REGION Network 36: STATE Num:120 StNextRdyInTransit
   RUNG wire#powerrail
      Contact( #sStNextRdyInTransit )
      wire#w1
      I_Contact( #sStWtResetRel )
      I_Contact( #sStNextRdyInTransit_T1 )
      I_Contact( #sStNextRdyInTransit_T2 )
      wire#w2
      Coil( #sStNextRdyInTransit )
   END_RUNG
   RUNG wire#powerrail
      Contact( #sStRecovery_T4 )
   END_RUNG wire#w1
   RUNG wire#powerrail
      Contact( #sStWtLifterAtPosn1_T1 )
   END_RUNG wire#w1
   RUNG wire#w2
      { S7_GenerateENO := "TRUE" } Move(in := 120, out1 => #StateNo)
   END_RUNG
   // the same network as SCL:
   #sStNextRdyInTransit := (#sStNextRdyInTransit OR #sStRecovery_T4 OR #sStWtLifterAtPosn1_T1) AND NOT #sStWtResetRel AND NOT #sStNextRdyInTransit_T1 AND NOT #sStNextRdyInTransit_T2;
   IF #sStNextRdyInTransit THEN #StateNo := 120; END_IF;
END_REGION

REGION Network 37: Transition for STATE Num:130 StNextRdyInTransit_1
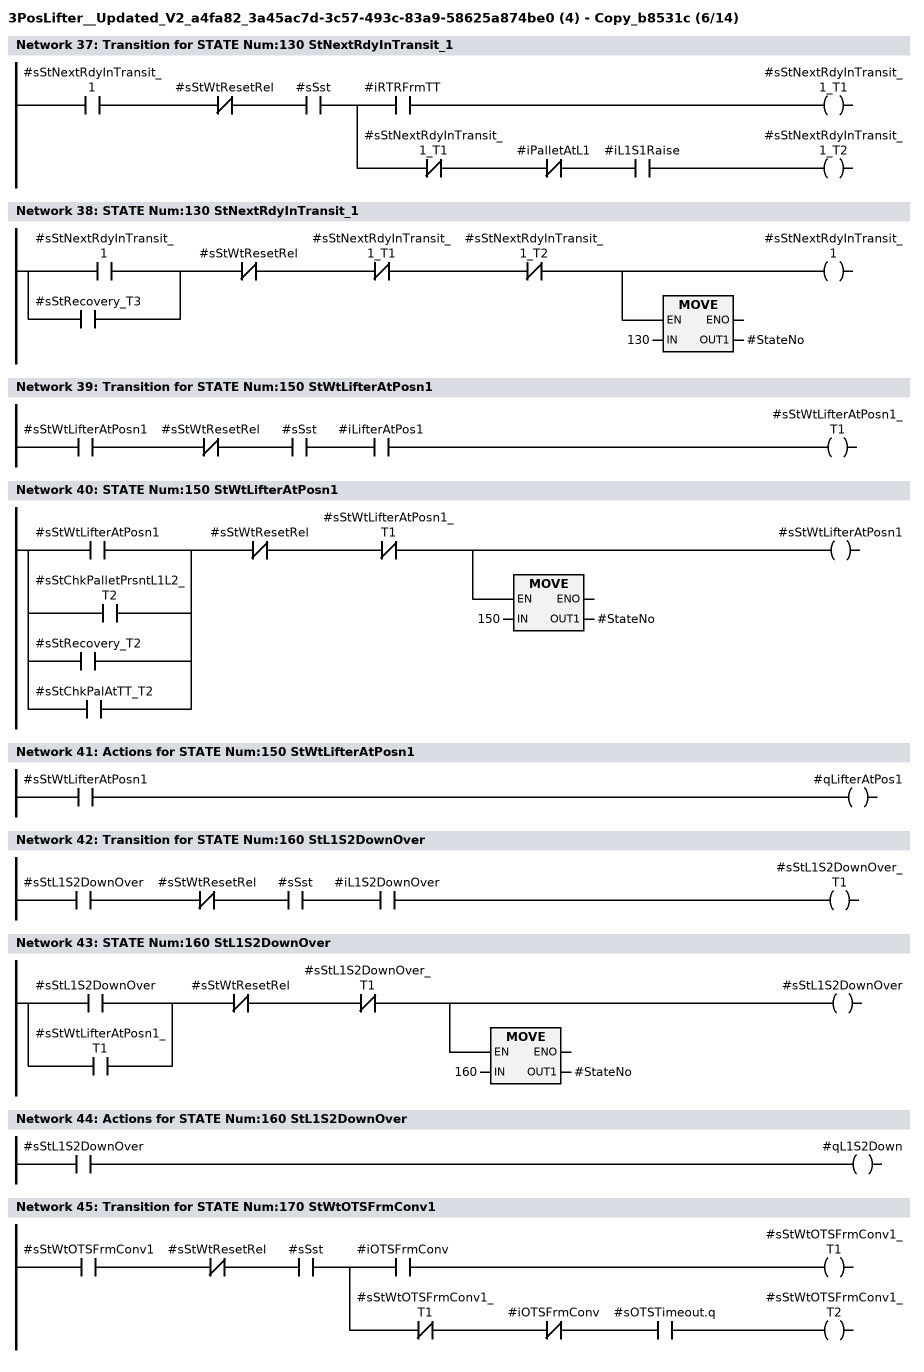
   RUNG wire#powerrail
      Contact( #sStNextRdyInTransit_1 )
      I_Contact( #sStWtResetRel )
      Contact( #sSst )
      wire#w1
      Contact( #iRTRFrmTT )
      Coil( #sStNextRdyInTransit_1_T1 )
   END_RUNG
   RUNG wire#w1
      I_Contact( #sStNextRdyInTransit_1_T1 )
      I_Contact( #iPalletAtL1 )
      Contact( #iL1S1Raise )
      Coil( #sStNextRdyInTransit_1_T2 )
   END_RUNG
   // the same network as SCL:
   #_w1 := #sStNextRdyInTransit_1 AND NOT #sStWtResetRel AND #sSst;
   #sStNextRdyInTransit_1_T1 := #_w1 AND #iRTRFrmTT;
   #sStNextRdyInTransit_1_T2 := #_w1 AND NOT #sStNextRdyInTransit_1_T1 AND NOT #iPalletAtL1 AND #iL1S1Raise;
END_REGION

REGION Network 38: STATE Num:130 StNextRdyInTransit_1
   RUNG wire#powerrail
      Contact( #sStNextRdyInTransit_1 )
      wire#w1
      I_Contact( #sStWtResetRel )
      I_Contact( #sStNextRdyInTransit_1_T1 )
      I_Contact( #sStNextRdyInTransit_1_T2 )
      wire#w2
      Coil( #sStNextRdyInTransit_1 )
   END_RUNG
   RUNG wire#powerrail
      Contact( #sStRecovery_T3 )
   END_RUNG wire#w1
   RUNG wire#w2
      { S7_GenerateENO := "TRUE" } Move(in := 130, out1 => #StateNo)
   END_RUNG
   // the same network as SCL:
   #sStNextRdyInTransit_1 := (#sStNextRdyInTransit_1 OR #sStRecovery_T3) AND NOT #sStWtResetRel AND NOT #sStNextRdyInTransit_1_T1 AND NOT #sStNextRdyInTransit_1_T2;
   IF #sStNextRdyInTransit_1 THEN #StateNo := 130; END_IF;
END_REGION

REGION Network 39: Transition for STATE Num:150 StWtLifterAtPosn1
   RUNG wire#powerrail
      Contact( #sStWtLifterAtPosn1 )
      I_Contact( #sStWtResetRel )
      Contact( #sSst )
      Contact( #iLifterAtPos1 )
      Coil( #sStWtLifterAtPosn1_T1 )
   END_RUNG
   // the same network as SCL:
   #sStWtLifterAtPosn1_T1 := #sStWtLifterAtPosn1 AND NOT #sStWtResetRel AND #sSst AND #iLifterAtPos1;
END_REGION

REGION Network 40: STATE Num:150 StWtLifterAtPosn1
   RUNG wire#powerrail
      Contact( #sStWtLifterAtPosn1 )
      wire#w1
      I_Contact( #sStWtResetRel )
      I_Contact( #sStWtLifterAtPosn1_T1 )
      wire#w2
      Coil( #sStWtLifterAtPosn1 )
   END_RUNG
   RUNG wire#powerrail
      Contact( #sStChkPalletPrsntL1L2_T2 )
   END_RUNG wire#w1
   RUNG wire#powerrail
      Contact( #sStRecovery_T2 )
   END_RUNG wire#w1
   RUNG wire#powerrail
      Contact( #sStChkPalAtTT_T2 )
   END_RUNG wire#w1
   RUNG wire#w2
      { S7_GenerateENO := "TRUE" } Move(in := 150, out1 => #StateNo)
   END_RUNG
   // the same network as SCL:
   #sStWtLifterAtPosn1 := (#sStWtLifterAtPosn1 OR #sStChkPalletPrsntL1L2_T2 OR #sStRecovery_T2 OR #sStChkPalAtTT_T2) AND NOT #sStWtResetRel AND NOT #sStWtLifterAtPosn1_T1;
   IF #sStWtLifterAtPosn1 THEN #StateNo := 150; END_IF;
END_REGION

REGION Network 41: Actions for STATE Num:150 StWtLifterAtPosn1
   RUNG wire#powerrail
      Contact( #sStWtLifterAtPosn1 )
      Coil( #qLifterAtPos1 )
   END_RUNG
   // the same network as SCL:
   #qLifterAtPos1 := #sStWtLifterAtPosn1;
END_REGION

REGION Network 42: Transition for STATE Num:160 StL1S2DownOver
   RUNG wire#powerrail
      Contact( #sStL1S2DownOver )
      I_Contact( #sStWtResetRel )
      Contact( #sSst )
      Contact( #iL1S2DownOver )
      Coil( #sStL1S2DownOver_T1 )
   END_RUNG
   // the same network as SCL:
   #sStL1S2DownOver_T1 := #sStL1S2DownOver AND NOT #sStWtResetRel AND #sSst AND #iL1S2DownOver;
END_REGION

REGION Network 43: STATE Num:160 StL1S2DownOver
   RUNG wire#powerrail
      Contact( #sStL1S2DownOver )
      wire#w1
      I_Contact( #sStWtResetRel )
      I_Contact( #sStL1S2DownOver_T1 )
      wire#w2
      Coil( #sStL1S2DownOver )
   END_RUNG
   RUNG wire#powerrail
      Contact( #sStWtLifterAtPosn1_T1 )
   END_RUNG wire#w1
   RUNG wire#w2
      { S7_GenerateENO := "TRUE" } Move(in := 160, out1 => #StateNo)
   END_RUNG
   // the same network as SCL:
   #sStL1S2DownOver := (#sStL1S2DownOver OR #sStWtLifterAtPosn1_T1) AND NOT #sStWtResetRel AND NOT #sStL1S2DownOver_T1;
   IF #sStL1S2DownOver THEN #StateNo := 160; END_IF;
END_REGION

REGION Network 44: Actions for STATE Num:160 StL1S2DownOver
   RUNG wire#powerrail
      Contact( #sStL1S2DownOver )
      Coil( #qL1S2Down )
   END_RUNG
   // the same network as SCL:
   #qL1S2Down := #sStL1S2DownOver;
END_REGION

REGION Network 45: Transition for STATE Num:170 StWtOTSFrmConv1
   RUNG wire#powerrail
      Contact( #sStWtOTSFrmConv1 )
      I_Contact( #sStWtResetRel )
      Contact( #sSst )
      wire#w1
      Contact( #iOTSFrmConv )
      Coil( #sStWtOTSFrmConv1_T1 )
   END_RUNG
   RUNG wire#w1
      I_Contact( #sStWtOTSFrmConv1_T1 )
      I_Contact( #iOTSFrmConv )
      Contact( #sOTSTimeout.q )
      Coil( #sStWtOTSFrmConv1_T2 )
   END_RUNG
   // the same network as SCL:
   #_w1 := #sStWtOTSFrmConv1 AND NOT #sStWtResetRel AND #sSst;
   #sStWtOTSFrmConv1_T1 := #_w1 AND #iOTSFrmConv;
   #sStWtOTSFrmConv1_T2 := #_w1 AND NOT #sStWtOTSFrmConv1_T1 AND NOT #iOTSFrmConv AND #sOTSTimeout.q;
END_REGION

REGION Network 46: STATE Num:170 StWtOTSFrmConv1
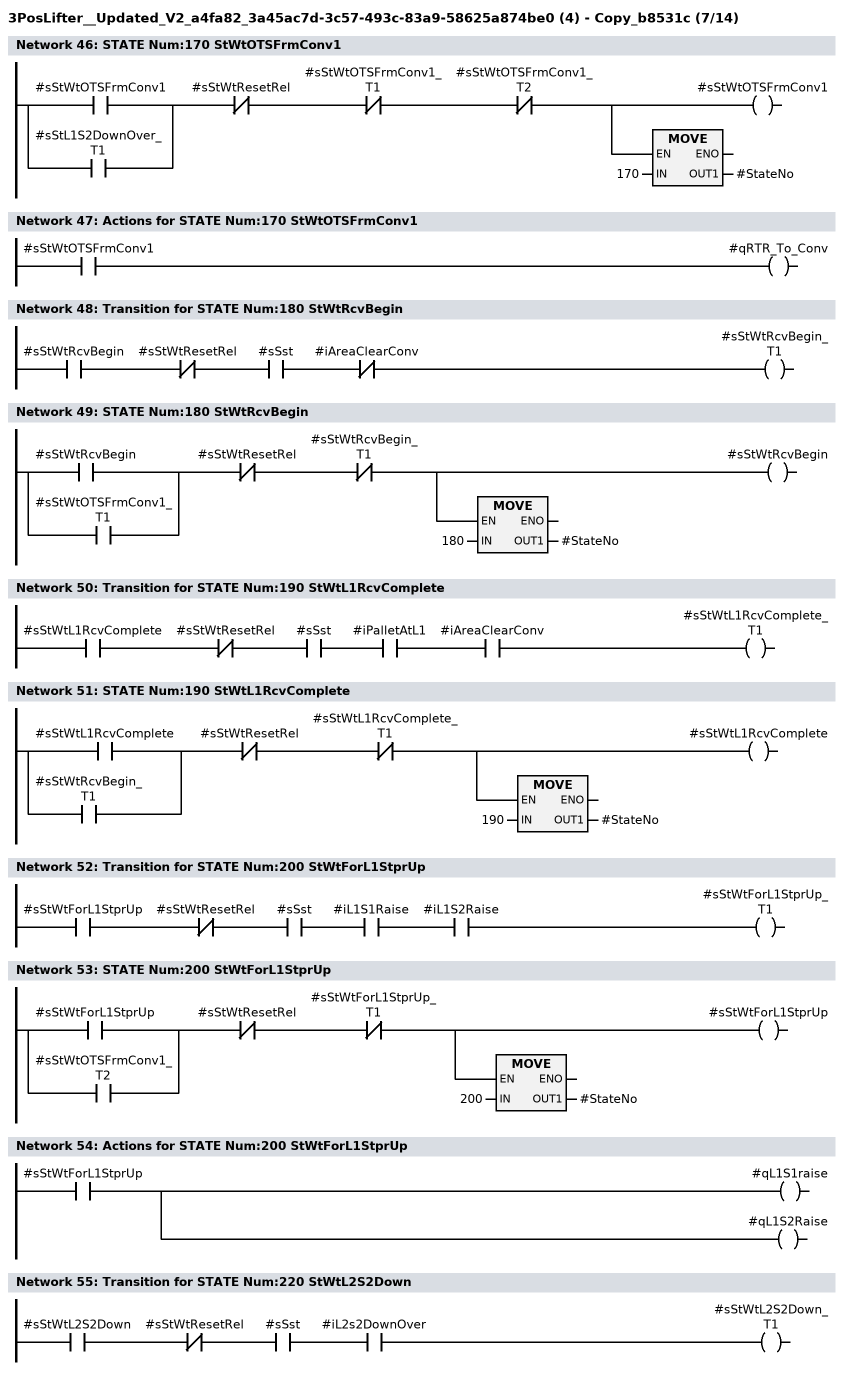
   RUNG wire#powerrail
      Contact( #sStWtOTSFrmConv1 )
      wire#w1
      I_Contact( #sStWtResetRel )
      I_Contact( #sStWtOTSFrmConv1_T1 )
      I_Contact( #sStWtOTSFrmConv1_T2 )
      wire#w2
      Coil( #sStWtOTSFrmConv1 )
   END_RUNG
   RUNG wire#powerrail
      Contact( #sStL1S2DownOver_T1 )
   END_RUNG wire#w1
   RUNG wire#w2
      { S7_GenerateENO := "TRUE" } Move(in := 170, out1 => #StateNo)
   END_RUNG
   // the same network as SCL:
   #sStWtOTSFrmConv1 := (#sStWtOTSFrmConv1 OR #sStL1S2DownOver_T1) AND NOT #sStWtResetRel AND NOT #sStWtOTSFrmConv1_T1 AND NOT #sStWtOTSFrmConv1_T2;
   IF #sStWtOTSFrmConv1 THEN #StateNo := 170; END_IF;
END_REGION

REGION Network 47: Actions for STATE Num:170 StWtOTSFrmConv1
   RUNG wire#powerrail
      Contact( #sStWtOTSFrmConv1 )
      Coil( #qRTR_To_Conv )
   END_RUNG
   // the same network as SCL:
   #qRTR_To_Conv := #sStWtOTSFrmConv1;
END_REGION

REGION Network 48: Transition for STATE Num:180 StWtRcvBegin
   RUNG wire#powerrail
      Contact( #sStWtRcvBegin )
      I_Contact( #sStWtResetRel )
      Contact( #sSst )
      I_Contact( #iAreaClearConv )
      Coil( #sStWtRcvBegin_T1 )
   END_RUNG
   // the same network as SCL:
   #sStWtRcvBegin_T1 := #sStWtRcvBegin AND NOT #sStWtResetRel AND #sSst AND NOT #iAreaClearConv;
END_REGION

REGION Network 49: STATE Num:180 StWtRcvBegin
   RUNG wire#powerrail
      Contact( #sStWtRcvBegin )
      wire#w1
      I_Contact( #sStWtResetRel )
      I_Contact( #sStWtRcvBegin_T1 )
      wire#w2
      Coil( #sStWtRcvBegin )
   END_RUNG
   RUNG wire#powerrail
      Contact( #sStWtOTSFrmConv1_T1 )
   END_RUNG wire#w1
   RUNG wire#w2
      { S7_GenerateENO := "TRUE" } Move(in := 180, out1 => #StateNo)
   END_RUNG
   // the same network as SCL:
   #sStWtRcvBegin := (#sStWtRcvBegin OR #sStWtOTSFrmConv1_T1) AND NOT #sStWtResetRel AND NOT #sStWtRcvBegin_T1;
   IF #sStWtRcvBegin THEN #StateNo := 180; END_IF;
END_REGION

REGION Network 50: Transition for STATE Num:190 StWtL1RcvComplete
   RUNG wire#powerrail
      Contact( #sStWtL1RcvComplete )
      I_Contact( #sStWtResetRel )
      Contact( #sSst )
      Contact( #iPalletAtL1 )
      Contact( #iAreaClearConv )
      Coil( #sStWtL1RcvComplete_T1 )
   END_RUNG
   // the same network as SCL:
   #sStWtL1RcvComplete_T1 := #sStWtL1RcvComplete AND NOT #sStWtResetRel AND #sSst AND #iPalletAtL1 AND #iAreaClearConv;
END_REGION

REGION Network 51: STATE Num:190 StWtL1RcvComplete
   RUNG wire#powerrail
      Contact( #sStWtL1RcvComplete )
      wire#w1
      I_Contact( #sStWtResetRel )
      I_Contact( #sStWtL1RcvComplete_T1 )
      wire#w2
      Coil( #sStWtL1RcvComplete )
   END_RUNG
   RUNG wire#powerrail
      Contact( #sStWtRcvBegin_T1 )
   END_RUNG wire#w1
   RUNG wire#w2
      { S7_GenerateENO := "TRUE" } Move(in := 190, out1 => #StateNo)
   END_RUNG
   // the same network as SCL:
   #sStWtL1RcvComplete := (#sStWtL1RcvComplete OR #sStWtRcvBegin_T1) AND NOT #sStWtResetRel AND NOT #sStWtL1RcvComplete_T1;
   IF #sStWtL1RcvComplete THEN #StateNo := 190; END_IF;
END_REGION

REGION Network 52: Transition for STATE Num:200 StWtForL1StprUp
   RUNG wire#powerrail
      Contact( #sStWtForL1StprUp )
      I_Contact( #sStWtResetRel )
      Contact( #sSst )
      Contact( #iL1S1Raise )
      Contact( #iL1S2Raise )
      Coil( #sStWtForL1StprUp_T1 )
   END_RUNG
   // the same network as SCL:
   #sStWtForL1StprUp_T1 := #sStWtForL1StprUp AND NOT #sStWtResetRel AND #sSst AND #iL1S1Raise AND #iL1S2Raise;
END_REGION

REGION Network 53: STATE Num:200 StWtForL1StprUp
   RUNG wire#powerrail
      Contact( #sStWtForL1StprUp )
      wire#w1
      I_Contact( #sStWtResetRel )
      I_Contact( #sStWtForL1StprUp_T1 )
      wire#w2
      Coil( #sStWtForL1StprUp )
   END_RUNG
   RUNG wire#powerrail
      Contact( #sStWtOTSFrmConv1_T2 )
   END_RUNG wire#w1
   RUNG wire#w2
      { S7_GenerateENO := "TRUE" } Move(in := 200, out1 => #StateNo)
   END_RUNG
   // the same network as SCL:
   #sStWtForL1StprUp := (#sStWtForL1StprUp OR #sStWtOTSFrmConv1_T2) AND NOT #sStWtResetRel AND NOT #sStWtForL1StprUp_T1;
   IF #sStWtForL1StprUp THEN #StateNo := 200; END_IF;
END_REGION

REGION Network 54: Actions for STATE Num:200 StWtForL1StprUp
   RUNG wire#powerrail
      Contact( #sStWtForL1StprUp )
      wire#w1
      Coil( #qL1S1raise )
   END_RUNG
   RUNG wire#w1
      Coil( #qL1S2Raise )
   END_RUNG
   // the same network as SCL:
   #qL1S1raise := #sStWtForL1StprUp;
   #qL1S2Raise := #sStWtForL1StprUp;
END_REGION

REGION Network 55: Transition for STATE Num:220 StWtL2S2Down
   RUNG wire#powerrail
      Contact( #sStWtL2S2Down )
      I_Contact( #sStWtResetRel )
      Contact( #sSst )
      Contact( #iL2s2DownOver )
      Coil( #sStWtL2S2Down_T1 )
   END_RUNG
   // the same network as SCL:
   #sStWtL2S2Down_T1 := #sStWtL2S2Down AND NOT #sStWtResetRel AND #sSst AND #iL2s2DownOver;
END_REGION

REGION Network 56: STATE Num:220 StWtL2S2Down
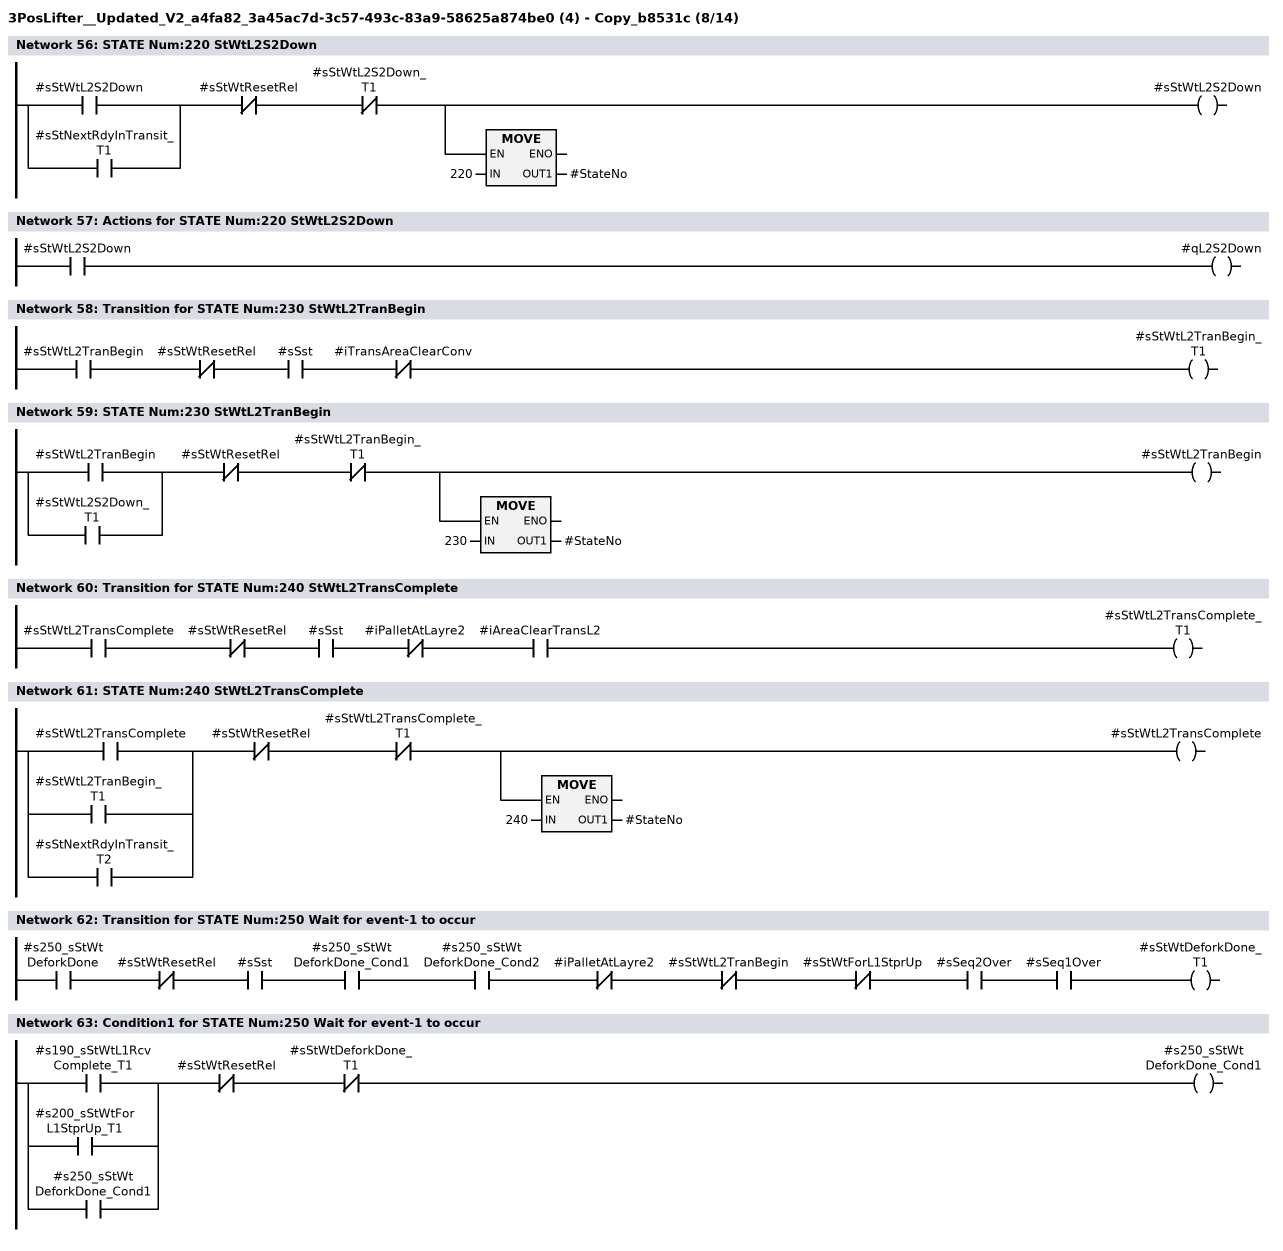
   RUNG wire#powerrail
      Contact( #sStWtL2S2Down )
      wire#w1
      I_Contact( #sStWtResetRel )
      I_Contact( #sStWtL2S2Down_T1 )
      wire#w2
      Coil( #sStWtL2S2Down )
   END_RUNG
   RUNG wire#powerrail
      Contact( #sStNextRdyInTransit_T1 )
   END_RUNG wire#w1
   RUNG wire#w2
      { S7_GenerateENO := "TRUE" } Move(in := 220, out1 => #StateNo)
   END_RUNG
   // the same network as SCL:
   #sStWtL2S2Down := (#sStWtL2S2Down OR #sStNextRdyInTransit_T1) AND NOT #sStWtResetRel AND NOT #sStWtL2S2Down_T1;
   IF #sStWtL2S2Down THEN #StateNo := 220; END_IF;
END_REGION

REGION Network 57: Actions for STATE Num:220 StWtL2S2Down
   RUNG wire#powerrail
      Contact( #sStWtL2S2Down )
      Coil( #qL2S2Down )
   END_RUNG
   // the same network as SCL:
   #qL2S2Down := #sStWtL2S2Down;
END_REGION

REGION Network 58: Transition for STATE Num:230 StWtL2TranBegin
   RUNG wire#powerrail
      Contact( #sStWtL2TranBegin )
      I_Contact( #sStWtResetRel )
      Contact( #sSst )
      I_Contact( #iTransAreaClearConv )
      Coil( #sStWtL2TranBegin_T1 )
   END_RUNG
   // the same network as SCL:
   #sStWtL2TranBegin_T1 := #sStWtL2TranBegin AND NOT #sStWtResetRel AND #sSst AND NOT #iTransAreaClearConv;
END_REGION

REGION Network 59: STATE Num:230 StWtL2TranBegin
   RUNG wire#powerrail
      Contact( #sStWtL2TranBegin )
      wire#w1
      I_Contact( #sStWtResetRel )
      I_Contact( #sStWtL2TranBegin_T1 )
      wire#w2
      Coil( #sStWtL2TranBegin )
   END_RUNG
   RUNG wire#powerrail
      Contact( #sStWtL2S2Down_T1 )
   END_RUNG wire#w1
   RUNG wire#w2
      { S7_GenerateENO := "TRUE" } Move(in := 230, out1 => #StateNo)
   END_RUNG
   // the same network as SCL:
   #sStWtL2TranBegin := (#sStWtL2TranBegin OR #sStWtL2S2Down_T1) AND NOT #sStWtResetRel AND NOT #sStWtL2TranBegin_T1;
   IF #sStWtL2TranBegin THEN #StateNo := 230; END_IF;
END_REGION

REGION Network 60: Transition for STATE Num:240 StWtL2TransComplete
   RUNG wire#powerrail
      Contact( #sStWtL2TransComplete )
      I_Contact( #sStWtResetRel )
      Contact( #sSst )
      I_Contact( #iPalletAtLayre2 )
      Contact( #iAreaClearTransL2 )
      Coil( #sStWtL2TransComplete_T1 )
   END_RUNG
   // the same network as SCL:
   #sStWtL2TransComplete_T1 := #sStWtL2TransComplete AND NOT #sStWtResetRel AND #sSst AND NOT #iPalletAtLayre2 AND #iAreaClearTransL2;
END_REGION

REGION Network 61: STATE Num:240 StWtL2TransComplete
   RUNG wire#powerrail
      Contact( #sStWtL2TransComplete )
      wire#w1
      I_Contact( #sStWtResetRel )
      I_Contact( #sStWtL2TransComplete_T1 )
      wire#w2
      Coil( #sStWtL2TransComplete )
   END_RUNG
   RUNG wire#powerrail
      Contact( #sStWtL2TranBegin_T1 )
   END_RUNG wire#w1
   RUNG wire#powerrail
      Contact( #sStNextRdyInTransit_T2 )
   END_RUNG wire#w1
   RUNG wire#w2
      { S7_GenerateENO := "TRUE" } Move(in := 240, out1 => #StateNo)
   END_RUNG
   // the same network as SCL:
   #sStWtL2TransComplete := (#sStWtL2TransComplete OR #sStWtL2TranBegin_T1 OR #sStNextRdyInTransit_T2) AND NOT #sStWtResetRel AND NOT #sStWtL2TransComplete_T1;
   IF #sStWtL2TransComplete THEN #StateNo := 240; END_IF;
END_REGION

REGION Network 62: Transition for STATE Num:250 Wait for event-1 to occur
   RUNG wire#powerrail
      Contact( #s250_sStWtDeforkDone )
      I_Contact( #sStWtResetRel )
      Contact( #sSst )
      Contact( #s250_sStWtDeforkDone_Cond1 )
      Contact( #s250_sStWtDeforkDone_Cond2 )
      I_Contact( #iPalletAtLayre2 )
      I_Contact( #sStWtL2TranBegin )
      I_Contact( #sStWtForL1StprUp )
      Contact( #sSeq2Over )
      Contact( #sSeq1Over )
      Coil( #sStWtDeforkDone_T1 )
   END_RUNG
   // the same network as SCL:
   #sStWtDeforkDone_T1 := #s250_sStWtDeforkDone AND NOT #sStWtResetRel AND #sSst AND #s250_sStWtDeforkDone_Cond1 AND #s250_sStWtDeforkDone_Cond2 AND NOT #iPalletAtLayre2 AND NOT #sStWtL2TranBegin AND NOT #sStWtForL1StprUp AND #sSeq2Over AND #sSeq1Over;
END_REGION

REGION Network 63: Condition1 for STATE Num:250 Wait for event-1 to occur
   RUNG wire#powerrail
      Contact( #s190_sStWtL1RcvComplete_T1 )
      wire#w1
      I_Contact( #sStWtResetRel )
      I_Contact( #sStWtDeforkDone_T1 )
      Coil( #s250_sStWtDeforkDone_Cond1 )
   END_RUNG
   RUNG wire#powerrail
      Contact( #s200_sStWtForL1StprUp_T1 )
   END_RUNG wire#w1
   RUNG wire#powerrail
      Contact( #s250_sStWtDeforkDone_Cond1 )
   END_RUNG wire#w1
   // the same network as SCL:
   #s250_sStWtDeforkDone_Cond1 := (#s190_sStWtL1RcvComplete_T1 OR #s200_sStWtForL1StprUp_T1 OR #s250_sStWtDeforkDone_Cond1) AND NOT #sStWtResetRel AND NOT #sStWtDeforkDone_T1;
END_REGION

REGION Network 64: Condition2 for STATE Num:250 Wait for event-1 to occur
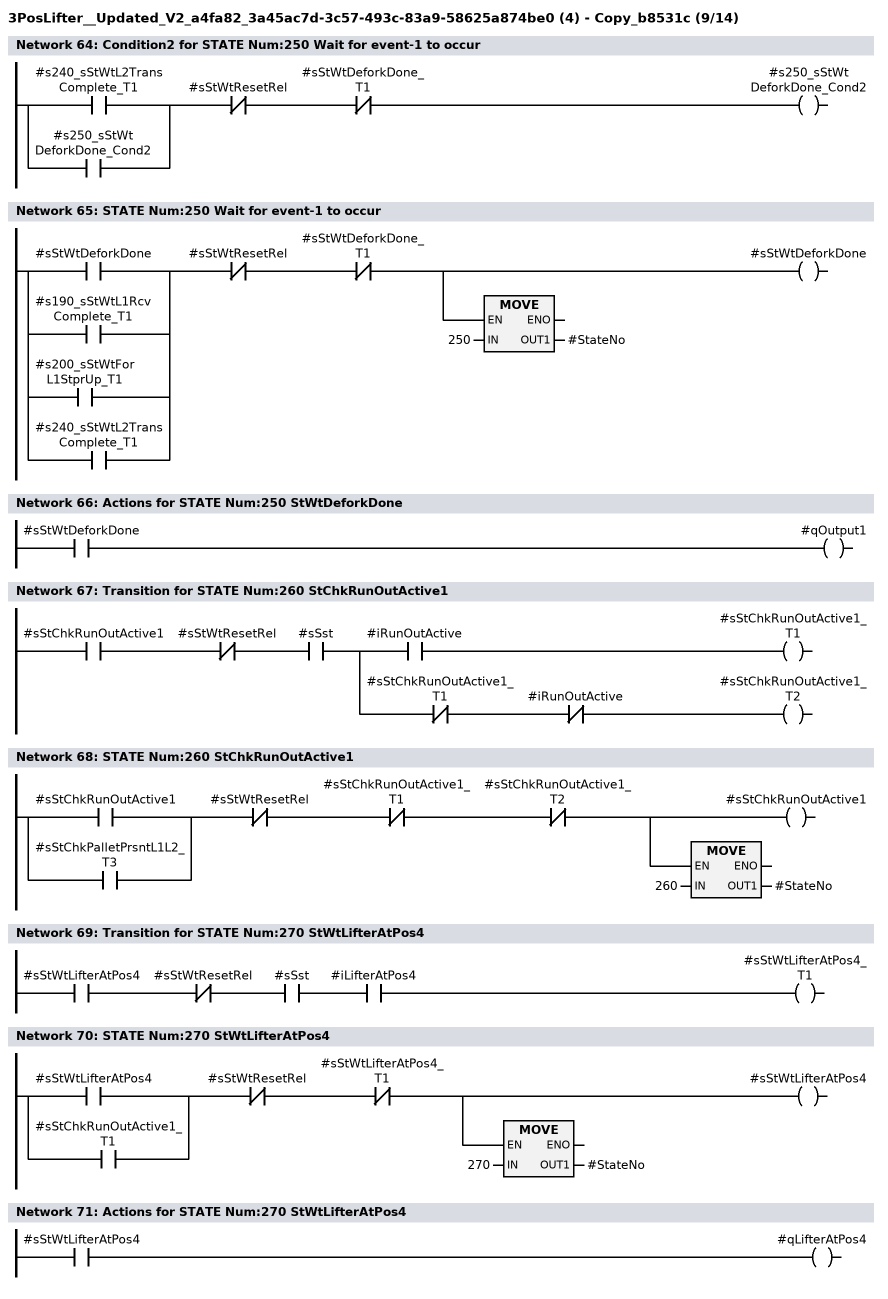
   RUNG wire#powerrail
      Contact( #s240_sStWtL2TransComplete_T1 )
      wire#w1
      I_Contact( #sStWtResetRel )
      I_Contact( #sStWtDeforkDone_T1 )
      Coil( #s250_sStWtDeforkDone_Cond2 )
   END_RUNG
   RUNG wire#powerrail
      Contact( #s250_sStWtDeforkDone_Cond2 )
   END_RUNG wire#w1
   // the same network as SCL:
   #s250_sStWtDeforkDone_Cond2 := (#s240_sStWtL2TransComplete_T1 OR #s250_sStWtDeforkDone_Cond2) AND NOT #sStWtResetRel AND NOT #sStWtDeforkDone_T1;
END_REGION

REGION Network 65: STATE Num:250 Wait for event-1 to occur
   RUNG wire#powerrail
      Contact( #sStWtDeforkDone )
      wire#w1
      I_Contact( #sStWtResetRel )
      I_Contact( #sStWtDeforkDone_T1 )
      wire#w2
      Coil( #sStWtDeforkDone )
   END_RUNG
   RUNG wire#powerrail
      Contact( #s190_sStWtL1RcvComplete_T1 )
   END_RUNG wire#w1
   RUNG wire#powerrail
      Contact( #s200_sStWtForL1StprUp_T1 )
   END_RUNG wire#w1
   RUNG wire#powerrail
      Contact( #s240_sStWtL2TransComplete_T1 )
   END_RUNG wire#w1
   RUNG wire#w2
      { S7_GenerateENO := "TRUE" } Move(in := 250, out1 => #StateNo)
   END_RUNG
   // the same network as SCL:
   #sStWtDeforkDone := (#sStWtDeforkDone OR #s190_sStWtL1RcvComplete_T1 OR #s200_sStWtForL1StprUp_T1 OR #s240_sStWtL2TransComplete_T1) AND NOT #sStWtResetRel AND NOT #sStWtDeforkDone_T1;
   IF #sStWtDeforkDone THEN #StateNo := 250; END_IF;
END_REGION

REGION Network 66: Actions for STATE Num:250 StWtDeforkDone
   RUNG wire#powerrail
      Contact( #sStWtDeforkDone )
      Coil( #qOutput1 )
   END_RUNG
   // the same network as SCL:
   #qOutput1 := #sStWtDeforkDone;
END_REGION

REGION Network 67: Transition for STATE Num:260 StChkRunOutActive1
   RUNG wire#powerrail
      Contact( #sStChkRunOutActive1 )
      I_Contact( #sStWtResetRel )
      Contact( #sSst )
      wire#w1
      Contact( #iRunOutActive )
      Coil( #sStChkRunOutActive1_T1 )
   END_RUNG
   RUNG wire#w1
      I_Contact( #sStChkRunOutActive1_T1 )
      I_Contact( #iRunOutActive )
      Coil( #sStChkRunOutActive1_T2 )
   END_RUNG
   // the same network as SCL:
   #_w1 := #sStChkRunOutActive1 AND NOT #sStWtResetRel AND #sSst;
   #sStChkRunOutActive1_T1 := #_w1 AND #iRunOutActive;
   #sStChkRunOutActive1_T2 := #_w1 AND NOT #sStChkRunOutActive1_T1 AND NOT #iRunOutActive;
END_REGION

REGION Network 68: STATE Num:260 StChkRunOutActive1
   RUNG wire#powerrail
      Contact( #sStChkRunOutActive1 )
      wire#w1
      I_Contact( #sStWtResetRel )
      I_Contact( #sStChkRunOutActive1_T1 )
      I_Contact( #sStChkRunOutActive1_T2 )
      wire#w2
      Coil( #sStChkRunOutActive1 )
   END_RUNG
   RUNG wire#powerrail
      Contact( #sStChkPalletPrsntL1L2_T3 )
   END_RUNG wire#w1
   RUNG wire#w2
      { S7_GenerateENO := "TRUE" } Move(in := 260, out1 => #StateNo)
   END_RUNG
   // the same network as SCL:
   #sStChkRunOutActive1 := (#sStChkRunOutActive1 OR #sStChkPalletPrsntL1L2_T3) AND NOT #sStWtResetRel AND NOT #sStChkRunOutActive1_T1 AND NOT #sStChkRunOutActive1_T2;
   IF #sStChkRunOutActive1 THEN #StateNo := 260; END_IF;
END_REGION

REGION Network 69: Transition for STATE Num:270 StWtLifterAtPos4
   RUNG wire#powerrail
      Contact( #sStWtLifterAtPos4 )
      I_Contact( #sStWtResetRel )
      Contact( #sSst )
      Contact( #iLifterAtPos4 )
      Coil( #sStWtLifterAtPos4_T1 )
   END_RUNG
   // the same network as SCL:
   #sStWtLifterAtPos4_T1 := #sStWtLifterAtPos4 AND NOT #sStWtResetRel AND #sSst AND #iLifterAtPos4;
END_REGION

REGION Network 70: STATE Num:270 StWtLifterAtPos4
   RUNG wire#powerrail
      Contact( #sStWtLifterAtPos4 )
      wire#w1
      I_Contact( #sStWtResetRel )
      I_Contact( #sStWtLifterAtPos4_T1 )
      wire#w2
      Coil( #sStWtLifterAtPos4 )
   END_RUNG
   RUNG wire#powerrail
      Contact( #sStChkRunOutActive1_T1 )
   END_RUNG wire#w1
   RUNG wire#w2
      { S7_GenerateENO := "TRUE" } Move(in := 270, out1 => #StateNo)
   END_RUNG
   // the same network as SCL:
   #sStWtLifterAtPos4 := (#sStWtLifterAtPos4 OR #sStChkRunOutActive1_T1) AND NOT #sStWtResetRel AND NOT #sStWtLifterAtPos4_T1;
   IF #sStWtLifterAtPos4 THEN #StateNo := 270; END_IF;
END_REGION

REGION Network 71: Actions for STATE Num:270 StWtLifterAtPos4
   RUNG wire#powerrail
      Contact( #sStWtLifterAtPos4 )
      Coil( #qLifterAtPos4 )
   END_RUNG
   // the same network as SCL:
   #qLifterAtPos4 := #sStWtLifterAtPos4;
END_REGION

REGION Network 72: Transition for STATE Num:280 StWtRTRFrmConvPos4
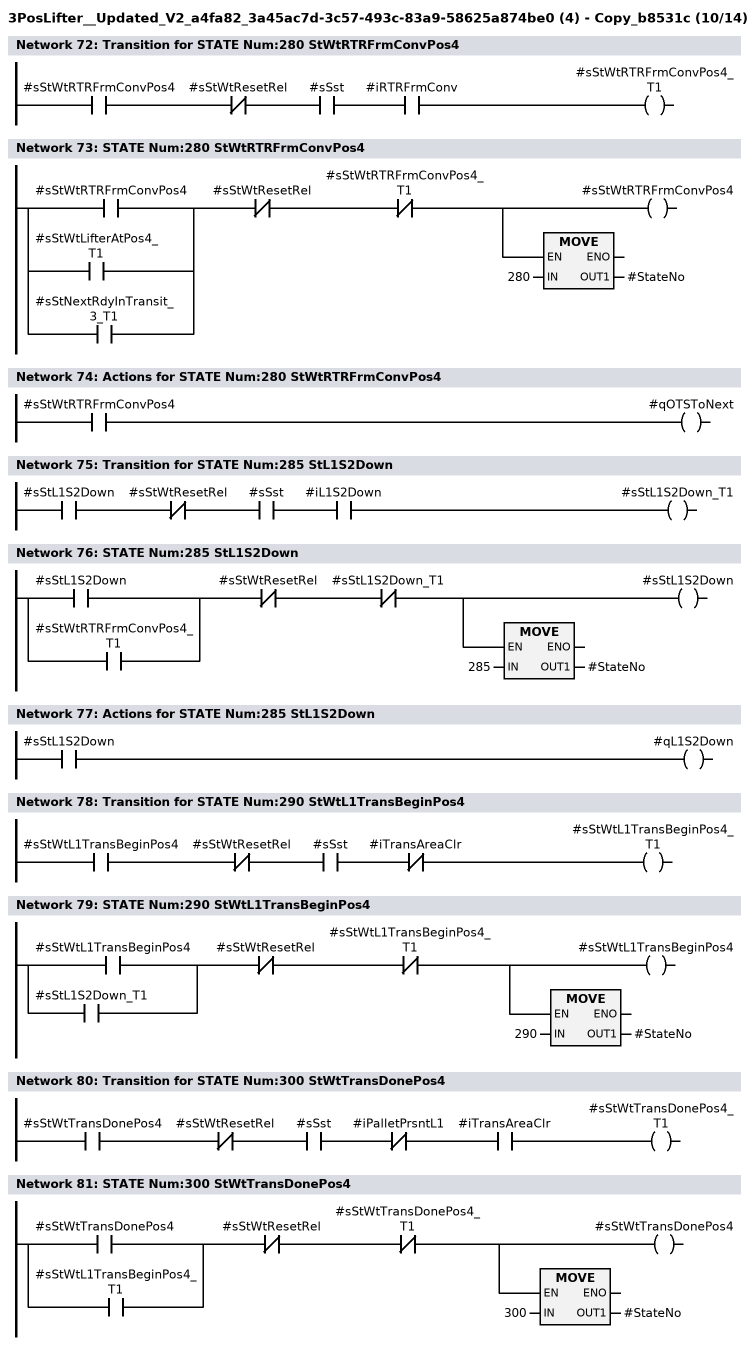
   RUNG wire#powerrail
      Contact( #sStWtRTRFrmConvPos4 )
      I_Contact( #sStWtResetRel )
      Contact( #sSst )
      Contact( #iRTRFrmConv )
      Coil( #sStWtRTRFrmConvPos4_T1 )
   END_RUNG
   // the same network as SCL:
   #sStWtRTRFrmConvPos4_T1 := #sStWtRTRFrmConvPos4 AND NOT #sStWtResetRel AND #sSst AND #iRTRFrmConv;
END_REGION

REGION Network 73: STATE Num:280 StWtRTRFrmConvPos4
   RUNG wire#powerrail
      Contact( #sStWtRTRFrmConvPos4 )
      wire#w1
      I_Contact( #sStWtResetRel )
      I_Contact( #sStWtRTRFrmConvPos4_T1 )
      wire#w2
      Coil( #sStWtRTRFrmConvPos4 )
   END_RUNG
   RUNG wire#powerrail
      Contact( #sStWtLifterAtPos4_T1 )
   END_RUNG wire#w1
   RUNG wire#powerrail
      Contact( #sStNextRdyInTransit_3_T1 )
   END_RUNG wire#w1
   RUNG wire#w2
      { S7_GenerateENO := "TRUE" } Move(in := 280, out1 => #StateNo)
   END_RUNG
   // the same network as SCL:
   #sStWtRTRFrmConvPos4 := (#sStWtRTRFrmConvPos4 OR #sStWtLifterAtPos4_T1 OR #sStNextRdyInTransit_3_T1) AND NOT #sStWtResetRel AND NOT #sStWtRTRFrmConvPos4_T1;
   IF #sStWtRTRFrmConvPos4 THEN #StateNo := 280; END_IF;
END_REGION

REGION Network 74: Actions for STATE Num:280 StWtRTRFrmConvPos4
   RUNG wire#powerrail
      Contact( #sStWtRTRFrmConvPos4 )
      Coil( #qOTSToNext )
   END_RUNG
   // the same network as SCL:
   #qOTSToNext := #sStWtRTRFrmConvPos4;
END_REGION

REGION Network 75: Transition for STATE Num:285 StL1S2Down
   RUNG wire#powerrail
      Contact( #sStL1S2Down )
      I_Contact( #sStWtResetRel )
      Contact( #sSst )
      Contact( #iL1S2Down )
      Coil( #sStL1S2Down_T1 )
   END_RUNG
   // the same network as SCL:
   #sStL1S2Down_T1 := #sStL1S2Down AND NOT #sStWtResetRel AND #sSst AND #iL1S2Down;
END_REGION

REGION Network 76: STATE Num:285 StL1S2Down
   RUNG wire#powerrail
      Contact( #sStL1S2Down )
      wire#w1
      I_Contact( #sStWtResetRel )
      I_Contact( #sStL1S2Down_T1 )
      wire#w2
      Coil( #sStL1S2Down )
   END_RUNG
   RUNG wire#powerrail
      Contact( #sStWtRTRFrmConvPos4_T1 )
   END_RUNG wire#w1
   RUNG wire#w2
      { S7_GenerateENO := "TRUE" } Move(in := 285, out1 => #StateNo)
   END_RUNG
   // the same network as SCL:
   #sStL1S2Down := (#sStL1S2Down OR #sStWtRTRFrmConvPos4_T1) AND NOT #sStWtResetRel AND NOT #sStL1S2Down_T1;
   IF #sStL1S2Down THEN #StateNo := 285; END_IF;
END_REGION

REGION Network 77: Actions for STATE Num:285 StL1S2Down
   RUNG wire#powerrail
      Contact( #sStL1S2Down )
      Coil( #qL1S2Down )
   END_RUNG
   // the same network as SCL:
   #qL1S2Down := #sStL1S2Down;
END_REGION

REGION Network 78: Transition for STATE Num:290 StWtL1TransBeginPos4
   RUNG wire#powerrail
      Contact( #sStWtL1TransBeginPos4 )
      I_Contact( #sStWtResetRel )
      Contact( #sSst )
      I_Contact( #iTransAreaClr )
      Coil( #sStWtL1TransBeginPos4_T1 )
   END_RUNG
   // the same network as SCL:
   #sStWtL1TransBeginPos4_T1 := #sStWtL1TransBeginPos4 AND NOT #sStWtResetRel AND #sSst AND NOT #iTransAreaClr;
END_REGION

REGION Network 79: STATE Num:290 StWtL1TransBeginPos4
   RUNG wire#powerrail
      Contact( #sStWtL1TransBeginPos4 )
      wire#w1
      I_Contact( #sStWtResetRel )
      I_Contact( #sStWtL1TransBeginPos4_T1 )
      wire#w2
      Coil( #sStWtL1TransBeginPos4 )
   END_RUNG
   RUNG wire#powerrail
      Contact( #sStL1S2Down_T1 )
   END_RUNG wire#w1
   RUNG wire#w2
      { S7_GenerateENO := "TRUE" } Move(in := 290, out1 => #StateNo)
   END_RUNG
   // the same network as SCL:
   #sStWtL1TransBeginPos4 := (#sStWtL1TransBeginPos4 OR #sStL1S2Down_T1) AND NOT #sStWtResetRel AND NOT #sStWtL1TransBeginPos4_T1;
   IF #sStWtL1TransBeginPos4 THEN #StateNo := 290; END_IF;
END_REGION

REGION Network 80: Transition for STATE Num:300 StWtTransDonePos4
   RUNG wire#powerrail
      Contact( #sStWtTransDonePos4 )
      I_Contact( #sStWtResetRel )
      Contact( #sSst )
      I_Contact( #iPalletPrsntL1 )
      Contact( #iTransAreaClr )
      Coil( #sStWtTransDonePos4_T1 )
   END_RUNG
   // the same network as SCL:
   #sStWtTransDonePos4_T1 := #sStWtTransDonePos4 AND NOT #sStWtResetRel AND #sSst AND NOT #iPalletPrsntL1 AND #iTransAreaClr;
END_REGION

REGION Network 81: STATE Num:300 StWtTransDonePos4
   RUNG wire#powerrail
      Contact( #sStWtTransDonePos4 )
      wire#w1
      I_Contact( #sStWtResetRel )
      I_Contact( #sStWtTransDonePos4_T1 )
      wire#w2
      Coil( #sStWtTransDonePos4 )
   END_RUNG
   RUNG wire#powerrail
      Contact( #sStWtL1TransBeginPos4_T1 )
   END_RUNG wire#w1
   RUNG wire#w2
      { S7_GenerateENO := "TRUE" } Move(in := 300, out1 => #StateNo)
   END_RUNG
   // the same network as SCL:
   #sStWtTransDonePos4 := (#sStWtTransDonePos4 OR #sStWtL1TransBeginPos4_T1) AND NOT #sStWtResetRel AND NOT #sStWtTransDonePos4_T1;
   IF #sStWtTransDonePos4 THEN #StateNo := 300; END_IF;
END_REGION

REGION Network 82: Transition for STATE Num:310 StChkPalletAtTT1
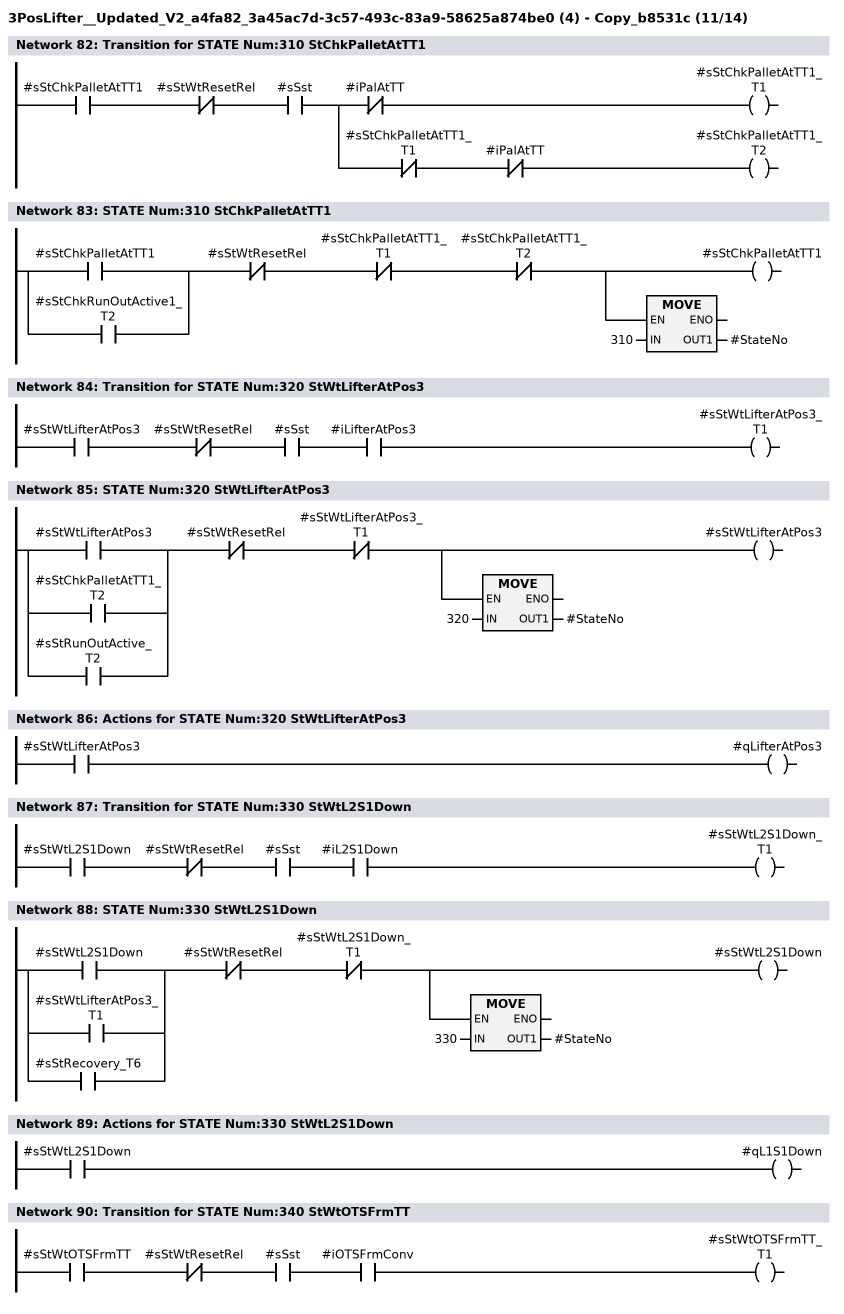
   RUNG wire#powerrail
      Contact( #sStChkPalletAtTT1 )
      I_Contact( #sStWtResetRel )
      Contact( #sSst )
      wire#w1
      I_Contact( #iPalAtTT )
      Coil( #sStChkPalletAtTT1_T1 )
   END_RUNG
   RUNG wire#w1
      I_Contact( #sStChkPalletAtTT1_T1 )
      I_Contact( #iPalAtTT )
      Coil( #sStChkPalletAtTT1_T2 )
   END_RUNG
   // the same network as SCL:
   #_w1 := #sStChkPalletAtTT1 AND NOT #sStWtResetRel AND #sSst;
   #sStChkPalletAtTT1_T1 := #_w1 AND NOT #iPalAtTT;
   #sStChkPalletAtTT1_T2 := #_w1 AND NOT #sStChkPalletAtTT1_T1 AND NOT #iPalAtTT;
END_REGION

REGION Network 83: STATE Num:310 StChkPalletAtTT1
   RUNG wire#powerrail
      Contact( #sStChkPalletAtTT1 )
      wire#w1
      I_Contact( #sStWtResetRel )
      I_Contact( #sStChkPalletAtTT1_T1 )
      I_Contact( #sStChkPalletAtTT1_T2 )
      wire#w2
      Coil( #sStChkPalletAtTT1 )
   END_RUNG
   RUNG wire#powerrail
      Contact( #sStChkRunOutActive1_T2 )
   END_RUNG wire#w1
   RUNG wire#w2
      { S7_GenerateENO := "TRUE" } Move(in := 310, out1 => #StateNo)
   END_RUNG
   // the same network as SCL:
   #sStChkPalletAtTT1 := (#sStChkPalletAtTT1 OR #sStChkRunOutActive1_T2) AND NOT #sStWtResetRel AND NOT #sStChkPalletAtTT1_T1 AND NOT #sStChkPalletAtTT1_T2;
   IF #sStChkPalletAtTT1 THEN #StateNo := 310; END_IF;
END_REGION

REGION Network 84: Transition for STATE Num:320 StWtLifterAtPos3
   RUNG wire#powerrail
      Contact( #sStWtLifterAtPos3 )
      I_Contact( #sStWtResetRel )
      Contact( #sSst )
      Contact( #iLifterAtPos3 )
      Coil( #sStWtLifterAtPos3_T1 )
   END_RUNG
   // the same network as SCL:
   #sStWtLifterAtPos3_T1 := #sStWtLifterAtPos3 AND NOT #sStWtResetRel AND #sSst AND #iLifterAtPos3;
END_REGION

REGION Network 85: STATE Num:320 StWtLifterAtPos3
   RUNG wire#powerrail
      Contact( #sStWtLifterAtPos3 )
      wire#w1
      I_Contact( #sStWtResetRel )
      I_Contact( #sStWtLifterAtPos3_T1 )
      wire#w2
      Coil( #sStWtLifterAtPos3 )
   END_RUNG
   RUNG wire#powerrail
      Contact( #sStChkPalletAtTT1_T2 )
   END_RUNG wire#w1
   RUNG wire#powerrail
      Contact( #sStRunOutActive_T2 )
   END_RUNG wire#w1
   RUNG wire#w2
      { S7_GenerateENO := "TRUE" } Move(in := 320, out1 => #StateNo)
   END_RUNG
   // the same network as SCL:
   #sStWtLifterAtPos3 := (#sStWtLifterAtPos3 OR #sStChkPalletAtTT1_T2 OR #sStRunOutActive_T2) AND NOT #sStWtResetRel AND NOT #sStWtLifterAtPos3_T1;
   IF #sStWtLifterAtPos3 THEN #StateNo := 320; END_IF;
END_REGION

REGION Network 86: Actions for STATE Num:320 StWtLifterAtPos3
   RUNG wire#powerrail
      Contact( #sStWtLifterAtPos3 )
      Coil( #qLifterAtPos3 )
   END_RUNG
   // the same network as SCL:
   #qLifterAtPos3 := #sStWtLifterAtPos3;
END_REGION

REGION Network 87: Transition for STATE Num:330 StWtL2S1Down
   RUNG wire#powerrail
      Contact( #sStWtL2S1Down )
      I_Contact( #sStWtResetRel )
      Contact( #sSst )
      Contact( #iL2S1Down )
      Coil( #sStWtL2S1Down_T1 )
   END_RUNG
   // the same network as SCL:
   #sStWtL2S1Down_T1 := #sStWtL2S1Down AND NOT #sStWtResetRel AND #sSst AND #iL2S1Down;
END_REGION

REGION Network 88: STATE Num:330 StWtL2S1Down
   RUNG wire#powerrail
      Contact( #sStWtL2S1Down )
      wire#w1
      I_Contact( #sStWtResetRel )
      I_Contact( #sStWtL2S1Down_T1 )
      wire#w2
      Coil( #sStWtL2S1Down )
   END_RUNG
   RUNG wire#powerrail
      Contact( #sStWtLifterAtPos3_T1 )
   END_RUNG wire#w1
   RUNG wire#powerrail
      Contact( #sStRecovery_T6 )
   END_RUNG wire#w1
   RUNG wire#w2
      { S7_GenerateENO := "TRUE" } Move(in := 330, out1 => #StateNo)
   END_RUNG
   // the same network as SCL:
   #sStWtL2S1Down := (#sStWtL2S1Down OR #sStWtLifterAtPos3_T1 OR #sStRecovery_T6) AND NOT #sStWtResetRel AND NOT #sStWtL2S1Down_T1;
   IF #sStWtL2S1Down THEN #StateNo := 330; END_IF;
END_REGION

REGION Network 89: Actions for STATE Num:330 StWtL2S1Down
   RUNG wire#powerrail
      Contact( #sStWtL2S1Down )
      Coil( #qL1S1Down )
   END_RUNG
   // the same network as SCL:
   #qL1S1Down := #sStWtL2S1Down;
END_REGION

REGION Network 90: Transition for STATE Num:340 StWtOTSFrmTT
   RUNG wire#powerrail
      Contact( #sStWtOTSFrmTT )
      I_Contact( #sStWtResetRel )
      Contact( #sSst )
      Contact( #iOTSFrmConv )
      Coil( #sStWtOTSFrmTT_T1 )
   END_RUNG
   // the same network as SCL:
   #sStWtOTSFrmTT_T1 := #sStWtOTSFrmTT AND NOT #sStWtResetRel AND #sSst AND #iOTSFrmConv;
END_REGION

REGION Network 91: STATE Num:340 StWtOTSFrmTT
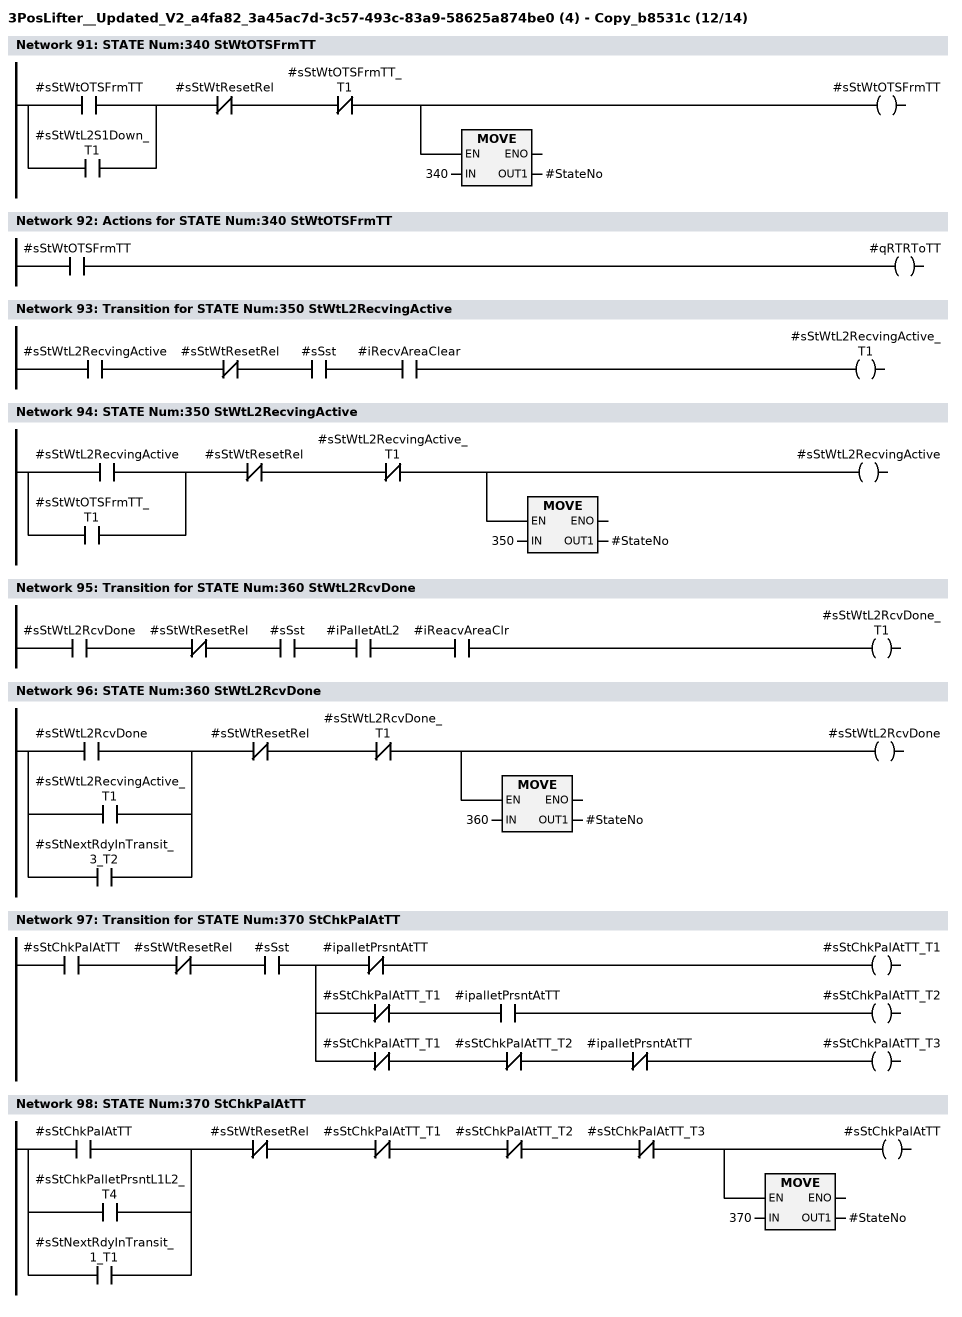
   RUNG wire#powerrail
      Contact( #sStWtOTSFrmTT )
      wire#w1
      I_Contact( #sStWtResetRel )
      I_Contact( #sStWtOTSFrmTT_T1 )
      wire#w2
      Coil( #sStWtOTSFrmTT )
   END_RUNG
   RUNG wire#powerrail
      Contact( #sStWtL2S1Down_T1 )
   END_RUNG wire#w1
   RUNG wire#w2
      { S7_GenerateENO := "TRUE" } Move(in := 340, out1 => #StateNo)
   END_RUNG
   // the same network as SCL:
   #sStWtOTSFrmTT := (#sStWtOTSFrmTT OR #sStWtL2S1Down_T1) AND NOT #sStWtResetRel AND NOT #sStWtOTSFrmTT_T1;
   IF #sStWtOTSFrmTT THEN #StateNo := 340; END_IF;
END_REGION

REGION Network 92: Actions for STATE Num:340 StWtOTSFrmTT
   RUNG wire#powerrail
      Contact( #sStWtOTSFrmTT )
      Coil( #qRTRToTT )
   END_RUNG
   // the same network as SCL:
   #qRTRToTT := #sStWtOTSFrmTT;
END_REGION

REGION Network 93: Transition for STATE Num:350 StWtL2RecvingActive
   RUNG wire#powerrail
      Contact( #sStWtL2RecvingActive )
      I_Contact( #sStWtResetRel )
      Contact( #sSst )
      Contact( #iRecvAreaClear )
      Coil( #sStWtL2RecvingActive_T1 )
   END_RUNG
   // the same network as SCL:
   #sStWtL2RecvingActive_T1 := #sStWtL2RecvingActive AND NOT #sStWtResetRel AND #sSst AND #iRecvAreaClear;
END_REGION

REGION Network 94: STATE Num:350 StWtL2RecvingActive
   RUNG wire#powerrail
      Contact( #sStWtL2RecvingActive )
      wire#w1
      I_Contact( #sStWtResetRel )
      I_Contact( #sStWtL2RecvingActive_T1 )
      wire#w2
      Coil( #sStWtL2RecvingActive )
   END_RUNG
   RUNG wire#powerrail
      Contact( #sStWtOTSFrmTT_T1 )
   END_RUNG wire#w1
   RUNG wire#w2
      { S7_GenerateENO := "TRUE" } Move(in := 350, out1 => #StateNo)
   END_RUNG
   // the same network as SCL:
   #sStWtL2RecvingActive := (#sStWtL2RecvingActive OR #sStWtOTSFrmTT_T1) AND NOT #sStWtResetRel AND NOT #sStWtL2RecvingActive_T1;
   IF #sStWtL2RecvingActive THEN #StateNo := 350; END_IF;
END_REGION

REGION Network 95: Transition for STATE Num:360 StWtL2RcvDone
   RUNG wire#powerrail
      Contact( #sStWtL2RcvDone )
      I_Contact( #sStWtResetRel )
      Contact( #sSst )
      Contact( #iPalletAtL2 )
      Contact( #iReacvAreaClr )
      Coil( #sStWtL2RcvDone_T1 )
   END_RUNG
   // the same network as SCL:
   #sStWtL2RcvDone_T1 := #sStWtL2RcvDone AND NOT #sStWtResetRel AND #sSst AND #iPalletAtL2 AND #iReacvAreaClr;
END_REGION

REGION Network 96: STATE Num:360 StWtL2RcvDone
   RUNG wire#powerrail
      Contact( #sStWtL2RcvDone )
      wire#w1
      I_Contact( #sStWtResetRel )
      I_Contact( #sStWtL2RcvDone_T1 )
      wire#w2
      Coil( #sStWtL2RcvDone )
   END_RUNG
   RUNG wire#powerrail
      Contact( #sStWtL2RecvingActive_T1 )
   END_RUNG wire#w1
   RUNG wire#powerrail
      Contact( #sStNextRdyInTransit_3_T2 )
   END_RUNG wire#w1
   RUNG wire#w2
      { S7_GenerateENO := "TRUE" } Move(in := 360, out1 => #StateNo)
   END_RUNG
   // the same network as SCL:
   #sStWtL2RcvDone := (#sStWtL2RcvDone OR #sStWtL2RecvingActive_T1 OR #sStNextRdyInTransit_3_T2) AND NOT #sStWtResetRel AND NOT #sStWtL2RcvDone_T1;
   IF #sStWtL2RcvDone THEN #StateNo := 360; END_IF;
END_REGION

REGION Network 97: Transition for STATE Num:370 StChkPalAtTT
   RUNG wire#powerrail
      Contact( #sStChkPalAtTT )
      I_Contact( #sStWtResetRel )
      Contact( #sSst )
      wire#w1
      I_Contact( #ipalletPrsntAtTT )
      Coil( #sStChkPalAtTT_T1 )
   END_RUNG
   RUNG wire#w1
      I_Contact( #sStChkPalAtTT_T1 )
      Contact( #ipalletPrsntAtTT )
      Coil( #sStChkPalAtTT_T2 )
   END_RUNG
   RUNG wire#w1
      I_Contact( #sStChkPalAtTT_T1 )
      I_Contact( #sStChkPalAtTT_T2 )
      I_Contact( #ipalletPrsntAtTT )
      Coil( #sStChkPalAtTT_T3 )
   END_RUNG
   // the same network as SCL:
   #_w1 := #sStChkPalAtTT AND NOT #sStWtResetRel AND #sSst;
   #sStChkPalAtTT_T1 := #_w1 AND NOT #ipalletPrsntAtTT;
   #sStChkPalAtTT_T2 := #_w1 AND NOT #sStChkPalAtTT_T1 AND #ipalletPrsntAtTT;
   #sStChkPalAtTT_T3 := #_w1 AND NOT #sStChkPalAtTT_T1 AND NOT #sStChkPalAtTT_T2 AND NOT #ipalletPrsntAtTT;
END_REGION

REGION Network 98: STATE Num:370 StChkPalAtTT
   RUNG wire#powerrail
      Contact( #sStChkPalAtTT )
      wire#w1
      I_Contact( #sStWtResetRel )
      I_Contact( #sStChkPalAtTT_T1 )
      I_Contact( #sStChkPalAtTT_T2 )
      I_Contact( #sStChkPalAtTT_T3 )
      wire#w2
      Coil( #sStChkPalAtTT )
   END_RUNG
   RUNG wire#powerrail
      Contact( #sStChkPalletPrsntL1L2_T4 )
   END_RUNG wire#w1
   RUNG wire#powerrail
      Contact( #sStNextRdyInTransit_1_T1 )
   END_RUNG wire#w1
   RUNG wire#w2
      { S7_GenerateENO := "TRUE" } Move(in := 370, out1 => #StateNo)
   END_RUNG
   // the same network as SCL:
   #sStChkPalAtTT := (#sStChkPalAtTT OR #sStChkPalletPrsntL1L2_T4 OR #sStNextRdyInTransit_1_T1) AND NOT #sStWtResetRel AND NOT #sStChkPalAtTT_T1 AND NOT #sStChkPalAtTT_T2 AND NOT #sStChkPalAtTT_T3;
   IF #sStChkPalAtTT THEN #StateNo := 370; END_IF;
END_REGION

REGION Network 99: Transition for STATE Num:380 StWtLifterAtPos2
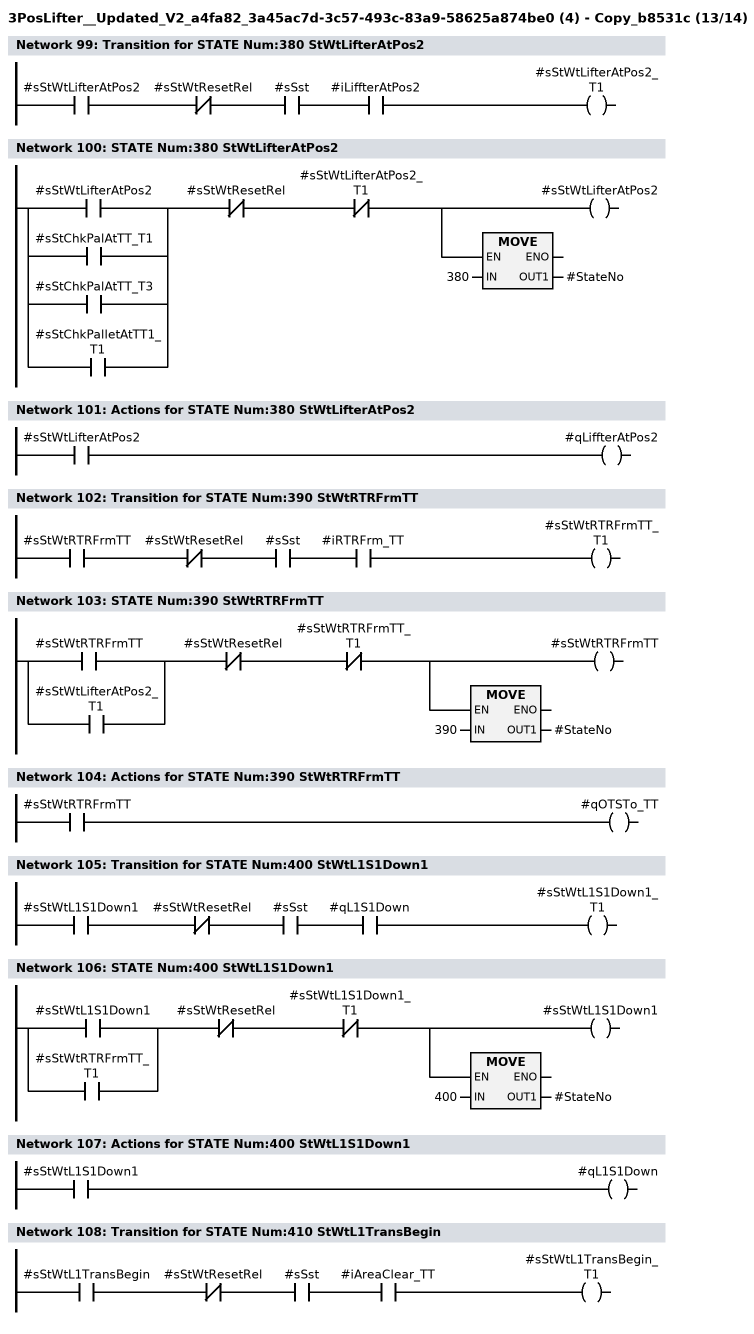
   RUNG wire#powerrail
      Contact( #sStWtLifterAtPos2 )
      I_Contact( #sStWtResetRel )
      Contact( #sSst )
      Contact( #iLiffterAtPos2 )
      Coil( #sStWtLifterAtPos2_T1 )
   END_RUNG
   // the same network as SCL:
   #sStWtLifterAtPos2_T1 := #sStWtLifterAtPos2 AND NOT #sStWtResetRel AND #sSst AND #iLiffterAtPos2;
END_REGION

REGION Network 100: STATE Num:380 StWtLifterAtPos2
   RUNG wire#powerrail
      Contact( #sStWtLifterAtPos2 )
      wire#w1
      I_Contact( #sStWtResetRel )
      I_Contact( #sStWtLifterAtPos2_T1 )
      wire#w2
      Coil( #sStWtLifterAtPos2 )
   END_RUNG
   RUNG wire#powerrail
      Contact( #sStChkPalAtTT_T1 )
   END_RUNG wire#w1
   RUNG wire#powerrail
      Contact( #sStChkPalAtTT_T3 )
   END_RUNG wire#w1
   RUNG wire#powerrail
      Contact( #sStChkPalletAtTT1_T1 )
   END_RUNG wire#w1
   RUNG wire#w2
      { S7_GenerateENO := "TRUE" } Move(in := 380, out1 => #StateNo)
   END_RUNG
   // the same network as SCL:
   #sStWtLifterAtPos2 := (#sStWtLifterAtPos2 OR #sStChkPalAtTT_T1 OR #sStChkPalAtTT_T3 OR #sStChkPalletAtTT1_T1) AND NOT #sStWtResetRel AND NOT #sStWtLifterAtPos2_T1;
   IF #sStWtLifterAtPos2 THEN #StateNo := 380; END_IF;
END_REGION

REGION Network 101: Actions for STATE Num:380 StWtLifterAtPos2
   RUNG wire#powerrail
      Contact( #sStWtLifterAtPos2 )
      Coil( #qLiffterAtPos2 )
   END_RUNG
   // the same network as SCL:
   #qLiffterAtPos2 := #sStWtLifterAtPos2;
END_REGION

REGION Network 102: Transition for STATE Num:390 StWtRTRFrmTT
   RUNG wire#powerrail
      Contact( #sStWtRTRFrmTT )
      I_Contact( #sStWtResetRel )
      Contact( #sSst )
      Contact( #iRTRFrm_TT )
      Coil( #sStWtRTRFrmTT_T1 )
   END_RUNG
   // the same network as SCL:
   #sStWtRTRFrmTT_T1 := #sStWtRTRFrmTT AND NOT #sStWtResetRel AND #sSst AND #iRTRFrm_TT;
END_REGION

REGION Network 103: STATE Num:390 StWtRTRFrmTT
   RUNG wire#powerrail
      Contact( #sStWtRTRFrmTT )
      wire#w1
      I_Contact( #sStWtResetRel )
      I_Contact( #sStWtRTRFrmTT_T1 )
      wire#w2
      Coil( #sStWtRTRFrmTT )
   END_RUNG
   RUNG wire#powerrail
      Contact( #sStWtLifterAtPos2_T1 )
   END_RUNG wire#w1
   RUNG wire#w2
      { S7_GenerateENO := "TRUE" } Move(in := 390, out1 => #StateNo)
   END_RUNG
   // the same network as SCL:
   #sStWtRTRFrmTT := (#sStWtRTRFrmTT OR #sStWtLifterAtPos2_T1) AND NOT #sStWtResetRel AND NOT #sStWtRTRFrmTT_T1;
   IF #sStWtRTRFrmTT THEN #StateNo := 390; END_IF;
END_REGION

REGION Network 104: Actions for STATE Num:390 StWtRTRFrmTT
   RUNG wire#powerrail
      Contact( #sStWtRTRFrmTT )
      Coil( #qOTSTo_TT )
   END_RUNG
   // the same network as SCL:
   #qOTSTo_TT := #sStWtRTRFrmTT;
END_REGION

REGION Network 105: Transition for STATE Num:400 StWtL1S1Down1
   RUNG wire#powerrail
      Contact( #sStWtL1S1Down1 )
      I_Contact( #sStWtResetRel )
      Contact( #sSst )
      Contact( #qL1S1Down )
      Coil( #sStWtL1S1Down1_T1 )
   END_RUNG
   // the same network as SCL:
   #sStWtL1S1Down1_T1 := #sStWtL1S1Down1 AND NOT #sStWtResetRel AND #sSst AND #qL1S1Down;
END_REGION

REGION Network 106: STATE Num:400 StWtL1S1Down1
   RUNG wire#powerrail
      Contact( #sStWtL1S1Down1 )
      wire#w1
      I_Contact( #sStWtResetRel )
      I_Contact( #sStWtL1S1Down1_T1 )
      wire#w2
      Coil( #sStWtL1S1Down1 )
   END_RUNG
   RUNG wire#powerrail
      Contact( #sStWtRTRFrmTT_T1 )
   END_RUNG wire#w1
   RUNG wire#w2
      { S7_GenerateENO := "TRUE" } Move(in := 400, out1 => #StateNo)
   END_RUNG
   // the same network as SCL:
   #sStWtL1S1Down1 := (#sStWtL1S1Down1 OR #sStWtRTRFrmTT_T1) AND NOT #sStWtResetRel AND NOT #sStWtL1S1Down1_T1;
   IF #sStWtL1S1Down1 THEN #StateNo := 400; END_IF;
END_REGION

REGION Network 107: Actions for STATE Num:400 StWtL1S1Down1
   RUNG wire#powerrail
      Contact( #sStWtL1S1Down1 )
      Coil( #qL1S1Down )
   END_RUNG
   // the same network as SCL:
   #qL1S1Down := #sStWtL1S1Down1;
END_REGION

REGION Network 108: Transition for STATE Num:410 StWtL1TransBegin
   RUNG wire#powerrail
      Contact( #sStWtL1TransBegin )
      I_Contact( #sStWtResetRel )
      Contact( #sSst )
      Contact( #iAreaClear_TT )
      Coil( #sStWtL1TransBegin_T1 )
   END_RUNG
   // the same network as SCL:
   #sStWtL1TransBegin_T1 := #sStWtL1TransBegin AND NOT #sStWtResetRel AND #sSst AND #iAreaClear_TT;
END_REGION

REGION Network 109: STATE Num:410 StWtL1TransBegin
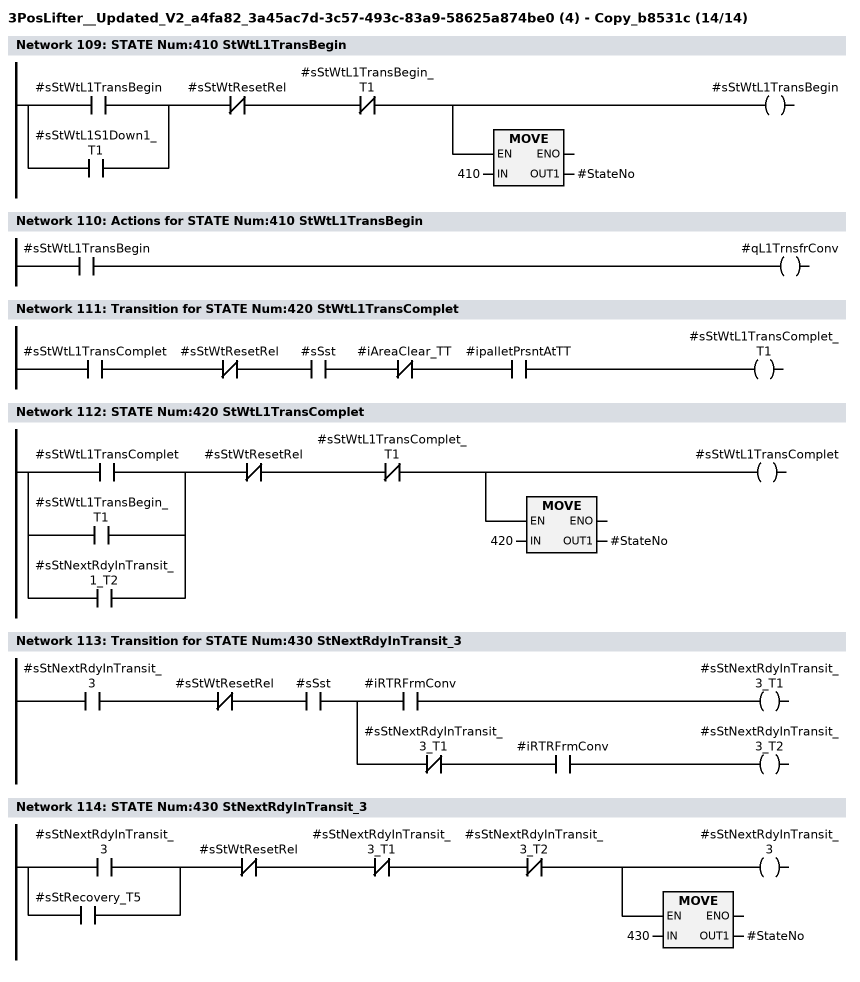
   RUNG wire#powerrail
      Contact( #sStWtL1TransBegin )
      wire#w1
      I_Contact( #sStWtResetRel )
      I_Contact( #sStWtL1TransBegin_T1 )
      wire#w2
      Coil( #sStWtL1TransBegin )
   END_RUNG
   RUNG wire#powerrail
      Contact( #sStWtL1S1Down1_T1 )
   END_RUNG wire#w1
   RUNG wire#w2
      { S7_GenerateENO := "TRUE" } Move(in := 410, out1 => #StateNo)
   END_RUNG
   // the same network as SCL:
   #sStWtL1TransBegin := (#sStWtL1TransBegin OR #sStWtL1S1Down1_T1) AND NOT #sStWtResetRel AND NOT #sStWtL1TransBegin_T1;
   IF #sStWtL1TransBegin THEN #StateNo := 410; END_IF;
END_REGION

REGION Network 110: Actions for STATE Num:410 StWtL1TransBegin
   RUNG wire#powerrail
      Contact( #sStWtL1TransBegin )
      Coil( #qL1TrnsfrConv )
   END_RUNG
   // the same network as SCL:
   #qL1TrnsfrConv := #sStWtL1TransBegin;
END_REGION

REGION Network 111: Transition for STATE Num:420 StWtL1TransComplet
   RUNG wire#powerrail
      Contact( #sStWtL1TransComplet )
      I_Contact( #sStWtResetRel )
      Contact( #sSst )
      I_Contact( #iAreaClear_TT )
      Contact( #ipalletPrsntAtTT )
      Coil( #sStWtL1TransComplet_T1 )
   END_RUNG
   // the same network as SCL:
   #sStWtL1TransComplet_T1 := #sStWtL1TransComplet AND NOT #sStWtResetRel AND #sSst AND NOT #iAreaClear_TT AND #ipalletPrsntAtTT;
END_REGION

REGION Network 112: STATE Num:420 StWtL1TransComplet
   RUNG wire#powerrail
      Contact( #sStWtL1TransComplet )
      wire#w1
      I_Contact( #sStWtResetRel )
      I_Contact( #sStWtL1TransComplet_T1 )
      wire#w2
      Coil( #sStWtL1TransComplet )
   END_RUNG
   RUNG wire#powerrail
      Contact( #sStWtL1TransBegin_T1 )
   END_RUNG wire#w1
   RUNG wire#powerrail
      Contact( #sStNextRdyInTransit_1_T2 )
   END_RUNG wire#w1
   RUNG wire#w2
      { S7_GenerateENO := "TRUE" } Move(in := 420, out1 => #StateNo)
   END_RUNG
   // the same network as SCL:
   #sStWtL1TransComplet := (#sStWtL1TransComplet OR #sStWtL1TransBegin_T1 OR #sStNextRdyInTransit_1_T2) AND NOT #sStWtResetRel AND NOT #sStWtL1TransComplet_T1;
   IF #sStWtL1TransComplet THEN #StateNo := 420; END_IF;
END_REGION

REGION Network 113: Transition for STATE Num:430 StNextRdyInTransit_3
   RUNG wire#powerrail
      Contact( #sStNextRdyInTransit_3 )
      I_Contact( #sStWtResetRel )
      Contact( #sSst )
      wire#w1
      Contact( #iRTRFrmConv )
      Coil( #sStNextRdyInTransit_3_T1 )
   END_RUNG
   RUNG wire#w1
      I_Contact( #sStNextRdyInTransit_3_T1 )
      Contact( #iRTRFrmConv )
      Coil( #sStNextRdyInTransit_3_T2 )
   END_RUNG
   // the same network as SCL:
   #_w1 := #sStNextRdyInTransit_3 AND NOT #sStWtResetRel AND #sSst;
   #sStNextRdyInTransit_3_T1 := #_w1 AND #iRTRFrmConv;
   #sStNextRdyInTransit_3_T2 := #_w1 AND NOT #sStNextRdyInTransit_3_T1 AND #iRTRFrmConv;
END_REGION

REGION Network 114: STATE Num:430 StNextRdyInTransit_3
   RUNG wire#powerrail
      Contact( #sStNextRdyInTransit_3 )
      wire#w1
      I_Contact( #sStWtResetRel )
      I_Contact( #sStNextRdyInTransit_3_T1 )
      I_Contact( #sStNextRdyInTransit_3_T2 )
      wire#w2
      Coil( #sStNextRdyInTransit_3 )
   END_RUNG
   RUNG wire#powerrail
      Contact( #sStRecovery_T5 )
   END_RUNG wire#w1
   RUNG wire#w2
      { S7_GenerateENO := "TRUE" } Move(in := 430, out1 => #StateNo)
   END_RUNG
   // the same network as SCL:
   #sStNextRdyInTransit_3 := (#sStNextRdyInTransit_3 OR #sStRecovery_T5) AND NOT #sStWtResetRel AND NOT #sStNextRdyInTransit_3_T1 AND NOT #sStNextRdyInTransit_3_T2;
   IF #sStNextRdyInTransit_3 THEN #StateNo := 430; END_IF;
END_REGION
END_FUNCTION_BLOCK

FUNCTION_BLOCK "S31808022001_Sequence_All_73b5c5_cfdfd9eb-ebd8-4267-a68e-df0ebcea3fa8 - Copy (2)_f93786"   // FB6, LAD
{ S7_Optimized_Access := 'TRUE' }
VERSION : 0.1
   VAR_INPUT
      iAutoRunning : Bool;
      iFaultReset : Bool;
      iOTS_Frm_Prev_TTDown : Bool;
      iOTS_Frm_Prev_TTUp : Bool;
      iPalletNtPrsntAtTTDown : Bool;
      iPalletNtPrsntAtTTUp : Bool;
      iPalletPrsnt_TTDown : Bool;
      iPalletPrsnt_TTUp : Bool;
      iPartReject : Bool;
      iRTR_Frm_Next_0DegTTUp : Bool;
      iRTR_Frm_Next_90DegTTUp : Bool;
      iRTR_Frm_Next_TTDown : Bool;
      iRecvAreaClr_TTDown : Bool;
      iRecvAreaClr_TTUp : Bool;
      iReset_fault : Bool;
      iRx_Frm_Prev_TTUp : Bool;
      iSstMode : Bool;
      iSstPB : Bool;
      iStprRaise_TTDown : Bool;
      iStprRaise_TTUp : Bool;
      iTTAt0Pos : Bool;
      iTTAt90Pos : Bool;
      iTTLocked : Bool;
      iTTUnlocked : Bool;
      iXferAreaClr_0DegTTDown : Bool;
      iXferAreaClr_0DegTTUp : Bool;
      iXferAreaClr_90DegTTUp : Bool;
   END_VAR
   VAR_OUTPUT
      qConvRun_TTDown : Bool;
      qConvRun_TTUp : Bool;
      qDelStprDown_TTUp : Bool;
      qOTS_Frm_TTDown : Bool;
      qOTS_Frm_TTUp : Bool;
      qOutput1 : Bool;
      qProcessStart : Bool;
      qRTR_Frm_TTDwn : Bool;
      qRTR_Frm_TTUp : Bool;
      qStprDown_TTDown : Bool;
      qStprDown_TTUp : Bool;
      qStprRaise_TTDown : Bool;
      qStprRaise_TTUp : Bool;
      qTTLockCmd : Bool;
      qTTUnlockCmd : Bool;
      qTT_0Deg : Bool;
      qTT_90Deg : Bool;
   END_VAR
   VAR_IN_OUT
      iqRX_Frn_Prev_TtDown : Bool;
      iqRx_Frm_Prev_TTUp : Bool;
      iqTx_To_Next_0DegTTDown : Bool;
      iqTx_To_Next_0DegTTUp : Bool;
      iqTx_To_Next_90DegTTUp : Bool;
   END_VAR
   VAR
      StateNo : Int;
      s100_StWtForTTUnlck : Bool;
      s100_StWtForTTUnlck_T1 : Bool;
      s10_StRecoveryCondition : Bool;
      s10_StRecoveryCondition_T1 : Bool;
      s10_StRecoveryCondition_T2 : Bool;
      s10_StRecoveryCondition_T3 : Bool;
      s10_StRecoveryCondition_T4 : Bool;
      s10_StRecoveryCondition_T5 : Bool;
      s10_StRecoveryCondition_T6 : Bool;
      s10_StRecoveryCondition_T7 : Bool;
      s110_StWtForTTTurn90 : Bool;
      s110_StWtForTTTurn90_T1 : Bool;
      s120_StWtForTTLck : Bool;
      s120_StWtForTTLck_T1 : Bool;
      s130_StChkTTDwnRdyToRecv : Bool;
      s130_StChkTTDwnRdyToRecv_T1 : Bool;
      s130_StChkTTDwnRdyToRecv_T2 : Bool;
      s140_StWtFrConveyorStrt : Bool;
      s140_StWtFrConveyorStrt_T1 : Bool;
      s150_StChkNxtStRdyToRecvTTUp : Bool;
      s150_StChkNxtStRdyToRecvTTUp_T1 : Bool;
      s150_StChkNxtStRdyToRecvTTUp_T2 : Bool;
      s15_StWaitForManCorrection : Bool;
      s15_StWaitForManCorrection_T1 : Bool;
      s160_StWtFrStprDn_CnvyrStrt : Bool;
      s160_StWtFrStprDn_CnvyrStrt_T1 : Bool;
      s165_StWtPalAbsnt : Bool;
      s165_StWtPalAbsnt_T1 : Bool;
      s167_StWtFrDeforkOvr : Bool;
      s167_StWtFrDeforkOvr_Cond1 : Bool;
      s167_StWtFrDeforkOvr_Cond2 : Bool;
      s167_StWtFrDeforkOvr_T1 : Bool;
      s170_StWtForTTUpStprUp : Bool;
      s170_StWtForTTUpStprUp_T1 : Bool;
      s180_StWtForTTUnlk : Bool;
      s180_StWtForTTUnlk_T1 : Bool;
      s190_StWtForTT_To_0 : Bool;
      s190_StWtForTT_To_0_T1 : Bool;
      s192_StWtForTTlok : Bool;
      s192_StWtForTTlok_T1 : Bool;
      s20_StChkForPalletPresent : Bool;
      s20_StChkForPalletPresent_T1 : Bool;
      s20_StChkForPalletPresent_T2 : Bool;
      s20_StChkForPalletPresent_T3 : Bool;
      s20_StChkForPalletPresent_T4 : Bool;
      s210_StWtFrTTUnlk : Bool;
      s210_StWtFrTTUnlk_T1 : Bool;
      s220_StWtFrTT_Trn_0 : Bool;
      s220_StWtFrTT_Trn_0_T1 : Bool;
      s230_StWtFrTTLock : Bool;
      s230_StWtFrTTLock_T1 : Bool;
      s240_StWtFRTRNxtStnTTDown : Bool;
      s240_StWtFRTRNxtStnTTDown_T1 : Bool;
      s240_StWtFRTRNxtStnTTDown_T2 : Bool;
      s250_StWtTTDnStprDn_CnvyrStr : Bool;
      s250_StWtTTDnStprDn_CnvyrStr_T1 : Bool;
      s260_StWtPalAbsent : Bool;
      s260_StWtPalAbsent_T1 : Bool;
      s270_StWtFrTTDwnStprUp : Bool;
      s270_StWtFrTTDwnStprUp_T1 : Bool;
      s280_StWtRFrOTSFRmPrev_TTUp : Bool;
      s280_StWtRFrOTSFRmPrev_TTUp_T1 : Bool;
      s290_StWtFrTTUpCnvyrStrt : Bool;
      s290_StWtFrTTUpCnvyrStrt_T1 : Bool;
      s300_StChkTTPos : Bool;
      s300_StChkTTPos_T1 : Bool;
      s300_StChkTTPos_T2 : Bool;
      s300_StChkTTPos_T3 : Bool;
      s30_StChckPartSts : Bool;
      s30_StChckPartSts_T1 : Bool;
      s310_StWtRTRFrmTTUpAt0 : Bool;
      s310_StWtRTRFrmTTUpAt0_T1 : Bool;
      s310_StWtRTRFrmTTUpAt0_T2 : Bool;
      s320_StWtFrTTUpCnvyrStrtAt0 : Bool;
      s320_StWtFrTTUpCnvyrStrtAt0_T1 : Bool;
      s340_StChkTTDwnRdyToRecvAt90 : Bool;
      s340_StChkTTDwnRdyToRecvAt90_T1 : Bool;
      s340_StChkTTDwnRdyToRecvAt90_T2 : Bool;
      s350_StWtCnvyrStrt90 : Bool;
      s350_StWtCnvyrStrt90_T1 : Bool;
      s365_StWtForTTUlkAtIbtwn : Bool;
      s365_StWtForTTUlkAtIbtwn_T1 : Bool;
      s370_StWtForTTTurnZrAtIbtwn : Bool;
      s370_StWtForTTTurnZrAtIbtwn_T1 : Bool;
      s380_StWtForTTLock : Bool;
      s380_StWtForTTLock_T1 : Bool;
      s400_StWt2Defork : Bool;
      s400_StWt2Defork_Cond1 : Bool;
      s400_StWt2Defork_Cond2 : Bool;
      s400_StWt2Defork_T1 : Bool;
      s40_StWtForTTUnlock : Bool;
      s40_StWtForTTUnlock_T1 : Bool;
      s410_StWtForTTUlkAtIbtwn : Bool;
      s410_StWtForTTUlkAtIbtwn_T1 : Bool;
      s415_StWtForTTTurn90AtIbtwn : Bool;
      s415_StWtForTTTurn90AtIbtwn_T1 : Bool;
      s420_StWtForTTLock1 : Bool;
      s420_StWtForTTLock1_T1 : Bool;
      s50_StWtForTTTurn0 : Bool;
      s50_StWtForTTTurn0_T1 : Bool;
      s60_StWtForTTLock : Bool;
      s60_StWtForTTLock_T1 : Bool;
      s70_StWtOTSfrmTTUp : Bool;
      s70_StWtOTSfrmTTUp_T1 : Bool;
      s80_StWtTTUpStpDwnCnvrStrt : Bool;
      s80_StWtTTUpStpDwnCnvrStrt_T1 : Bool;
      s85_StWtPalPresntAtRej : Bool;
      s85_StWtPalPresntAtRej_T1 : Bool;
      s90_StWtTTUpStprUp : Bool;
      s90_StWtTTUpStprUp_T1 : Bool;
      sDefork1Done : Bool;
      sDefork2Done : Bool;
      sOTSFrmDwnTout : Bool;
      sOTSFrmUpTout : Bool;
      sPalOnStop_TTDown : Bool;
      sPalOnStop_TTUp_0Deg : Bool;
      sPalOnStop_TTUp_90Deg : Bool;
      sPalletAbsnDebTTUp : Bool;
      sPalletAbsntDebTTDown : Bool;
      sPalletAbsntDebTTUp : Bool;
      sPalletPrsntDebTTDown : Bool;
      sPalletPrsntDebTTUp : Bool;
      sRTRFrmUpTout : Bool;
      sSst : Bool;
      sSstPulse : Bool;
      sSstRise : Bool;
      sStWtResetRel : Bool;
      sStWtResetRel_T1 : Bool;
      sTTDwnSeqOver : Bool;
      sTTDwn_0Pos_TX_Time : Bool;
      sTTDwn_90Pos_RX_Time : Bool;
      sTTDwn_Timer_ON : Bool;
      sTTUpSeqOver : Bool;
      sTTUp_90Pos_TX_Time : Bool;
      sTTUp_Timer_ON : Bool;
      sTrBothPalletPresent : Bool;
   END_VAR
   VAR_TEMP
      tOne : Bool;
   END_VAR
   VAR_TEMP   // added for the SCL form of the ladder/FBD networks
      _w1 : Bool;
   END_VAR
BEGIN

REGION Network 1
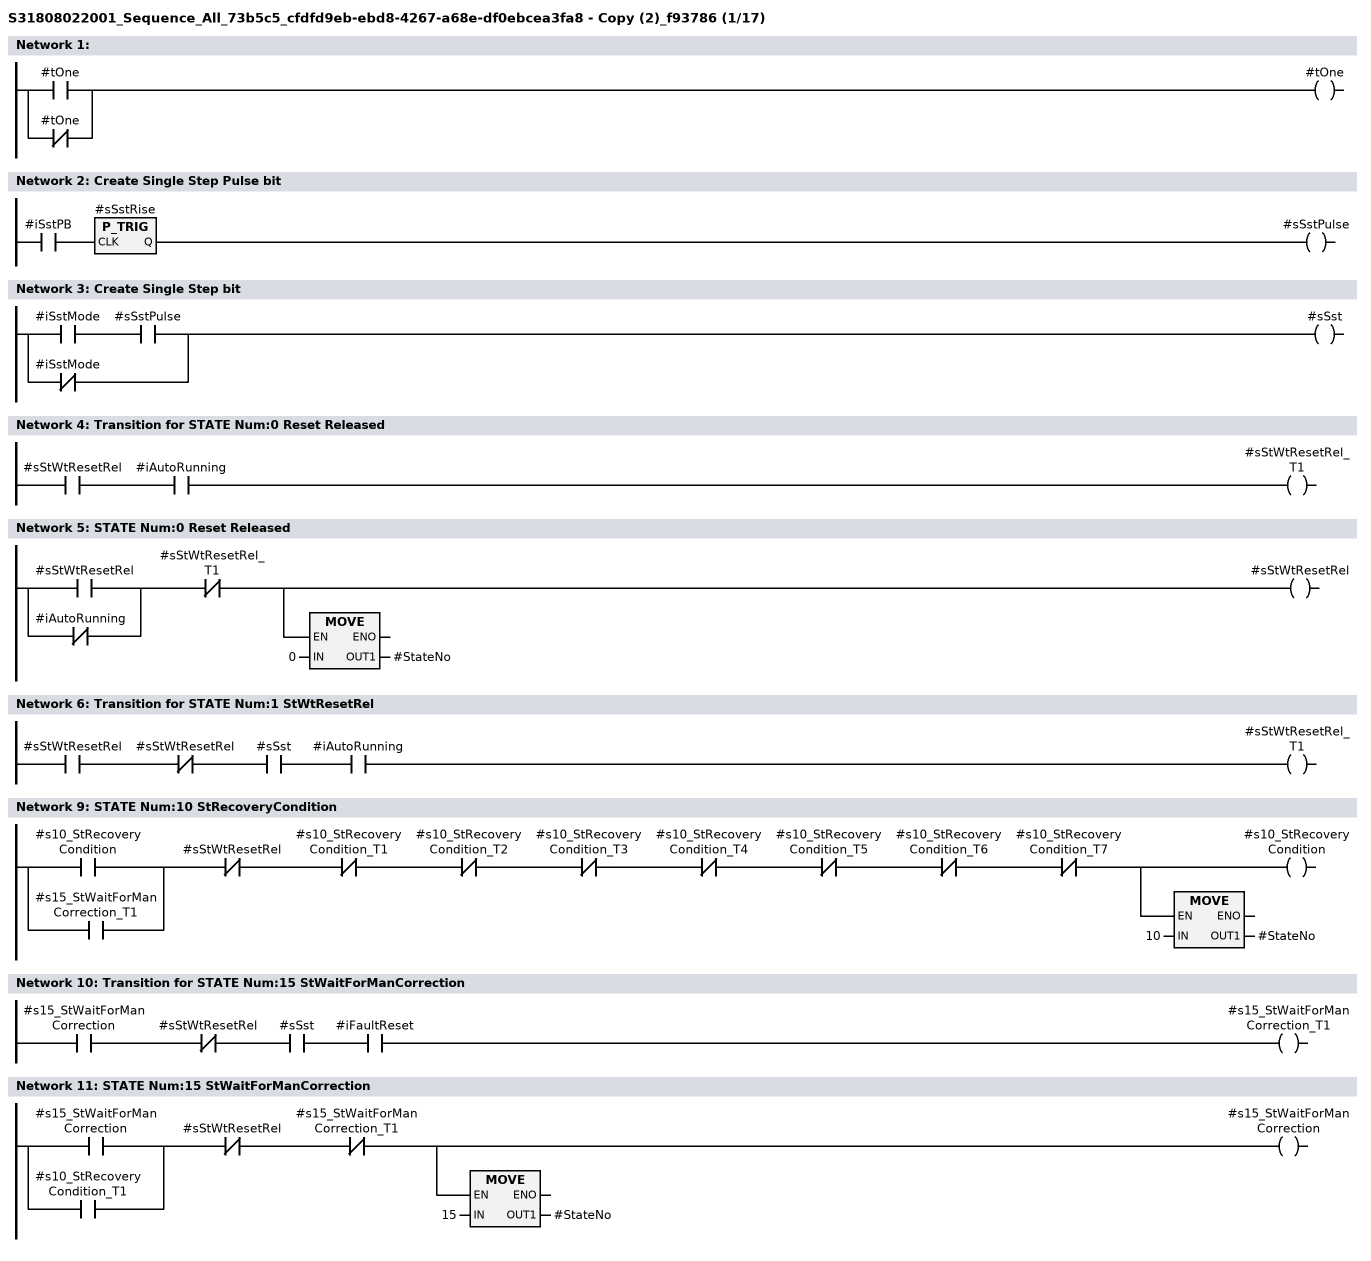
   RUNG wire#powerrail
      Contact( #tOne )
      wire#w1
      Coil( #tOne )
   END_RUNG
   RUNG wire#powerrail
      I_Contact( #tOne )
   END_RUNG wire#w1
   // the same network as SCL:
   #tOne := #tOne OR NOT #tOne;
END_REGION

REGION Network 2: Create Single Step Pulse bit
   RUNG wire#powerrail
      Contact( #iSstPB )
      P_Trig( #sSstRise )
      Coil( #sSstPulse )
   END_RUNG
   // the same network as SCL:
   #_w1 := #iSstPB AND NOT #sSstRise;   // rising edge
   #sSstRise := #iSstPB;
   #sSstPulse := #_w1;
END_REGION

REGION Network 3: Create Single Step bit
   RUNG wire#powerrail
      Contact( #iSstMode )
      Contact( #sSstPulse )
      wire#w1
      Coil( #sSst )
   END_RUNG
   RUNG wire#powerrail
      I_Contact( #iSstMode )
   END_RUNG wire#w1
   // the same network as SCL:
   #sSst := (#iSstMode AND #sSstPulse) OR NOT #iSstMode;
END_REGION

REGION Network 4: Transition for STATE Num:0 Reset Released
   RUNG wire#powerrail
      Contact( #sStWtResetRel )
      Contact( #iAutoRunning )
      Coil( #sStWtResetRel_T1 )
   END_RUNG
   // the same network as SCL:
   #sStWtResetRel_T1 := #sStWtResetRel AND #iAutoRunning;
END_REGION

REGION Network 5: STATE Num:0 Reset Released
   RUNG wire#powerrail
      Contact( #sStWtResetRel )
      wire#w1
      I_Contact( #sStWtResetRel_T1 )
      wire#w2
      Coil( #sStWtResetRel )
   END_RUNG
   RUNG wire#powerrail
      I_Contact( #iAutoRunning )
   END_RUNG wire#w1
   RUNG wire#w2
      { S7_GenerateENO := "TRUE" } Move(in := 0, out1 => #StateNo)
   END_RUNG
   // the same network as SCL:
   #sStWtResetRel := (#sStWtResetRel OR NOT #iAutoRunning) AND NOT #sStWtResetRel_T1;
   IF #sStWtResetRel THEN #StateNo := 0; END_IF;
END_REGION

REGION Network 6: Transition for STATE Num:1 StWtResetRel
   RUNG wire#powerrail
      Contact( #sStWtResetRel )
      I_Contact( #sStWtResetRel )
      Contact( #sSst )
      Contact( #iAutoRunning )
      Coil( #sStWtResetRel_T1 )
   END_RUNG
   // the same network as SCL:
   #sStWtResetRel_T1 := #sStWtResetRel AND NOT #sStWtResetRel AND #sSst AND #iAutoRunning;
END_REGION

REGION Network 7 (STL): STATE Num:1 StWtResetRel
         A(;
         O     #sStWtResetRel;
   //wrong transition variable removed
         );
         AN    #sStWtResetRel;
         AN    #sStWtResetRel_T1;
         =     <??.?>;
         A     <??.?>;
         BLD   102;
         =     #sStWtResetRel;
         A     <??.?>;
         JNB   Label_1;
         L     1;
         T     #StateNo;
   Label_1:NOP   0;
END_REGION

REGION Network 8 (STL): Transition for STATE Num:10 StRecoveryCondition
         A     #s10_StRecoveryCondition;
         AN    #sStWtResetRel;
         A     #sSst;
         =     <??.?>;
         A     <??.?>;
         A(;
         O(;
         A     #iRx_Frm_Prev_TTUp;
         AN    #iTTAt0Pos;
         );
         O(;
         A     #iqRX_Frn_Prev_TtDown;
         AN    #iTTAt90Pos;
         );
         O(;
         O     #iqTx_To_Next_90DegTTUp;
         O     #sPalOnStop_TTUp_90Deg;
         AN    #iTTAt90Pos;
         );
         O(;
         O     #iqTx_To_Next_0DegTTUp;
         O     #sPalOnStop_TTUp_0Deg;
         AN    #iTTAt0Pos;
         );
         O(;
         O     #iqTx_To_Next_0DegTTDown;
         O     #sPalOnStop_TTDown;
         AN    #iTTAt0Pos;
         );
         O(;
         O     #sPalOnStop_TTUp_0Deg;
         O     #sPalOnStop_TTUp_90Deg;
         O     #sPalOnStop_TTDown;
         A     #iTTUnlocked;
         );
         );
         =     #s10_StRecoveryCondition_T1;
         A     <??.?>;
         AN    #s10_StRecoveryCondition_T1;
         A(;
         O     #iqTx_To_Next_0DegTTUp;
         O     #sPalOnStop_TTUp_0Deg;
         );
         A     #iTTAt0Pos;
         A     #iTTLocked;
         =     #s10_StRecoveryCondition_T2;
         A     <??.?>;
         AN    #s10_StRecoveryCondition_T1;
         AN    #s10_StRecoveryCondition_T2;
         A(;
         O     #iqTx_To_Next_90DegTTUp;
         O     #sPalOnStop_TTUp_90Deg;
         );
         A     #iTTAt90Pos;
         A     #iTTLocked;
         =     #s10_StRecoveryCondition_T3;
         A     <??.?>;
         AN    #s10_StRecoveryCondition_T1;
         AN    #s10_StRecoveryCondition_T2;
         AN    #s10_StRecoveryCondition_T3;
         A(;
         O     #iqTx_To_Next_0DegTTDown;
         O     #sPalOnStop_TTDown;
         );
         A     #iTTAt0Pos;
         A     #iTTLocked;
         =     #s10_StRecoveryCondition_T4;
         A     <??.?>;
         AN    #s10_StRecoveryCondition_T1;
         AN    #s10_StRecoveryCondition_T2;
         AN    #s10_StRecoveryCondition_T3;
         AN    #s10_StRecoveryCondition_T4;
         A(;
         O     #iRx_Frm_Prev_TTUp;
         O     #iRecvAreaClr_TTUp;
         );
         A     #iTTAt0Pos;
         A     #iTTLocked;
         =     #s10_StRecoveryCondition_T5;
         A     <??.?>;
         AN    #s10_StRecoveryCondition_T1;
         AN    #s10_StRecoveryCondition_T2;
         AN    #s10_StRecoveryCondition_T3;
         AN    #s10_StRecoveryCondition_T4;
         AN    #s10_StRecoveryCondition_T5;
         A(;
         O     #iqRX_Frn_Prev_TtDown;
         ON    #iRecvAreaClr_TTDown;
         );
         A     #iTTAt90Pos;
         A     #iTTLocked;
         =     #s10_StRecoveryCondition_T6;
         A     <??.?>;
         AN    #s10_StRecoveryCondition_T1;
         AN    #s10_StRecoveryCondition_T2;
         AN    #s10_StRecoveryCondition_T3;
         AN    #s10_StRecoveryCondition_T4;
         AN    #s10_StRecoveryCondition_T5;
         AN    #s10_StRecoveryCondition_T6;
         A(;
         A(;
         A     #iXferAreaClr_90DegTTUp;
         A     #iXferAreaClr_0DegTTDown;
         A     #iRecvAreaClr_TTDown;
         A     #iRecvAreaClr_TTUp;
         );
         O(;
         AN    #sPalOnStop_TTUp_0Deg;
         AN    #sPalOnStop_TTUp_90Deg;
         AN    #sPalOnStop_TTDown;
         );
         O(;
         AN    #iqTx_To_Next_90DegTTUp;
         AN    #iqTx_To_Next_0DegTTUp;
         AN    #iqTx_To_Next_0DegTTDown;
         AN    #iqRX_Frn_Prev_TtDown;
         AN    #iRx_Frm_Prev_TTUp;
         );
         );
         =     #s10_StRecoveryCondition_T7;
END_REGION

REGION Network 9: STATE Num:10 StRecoveryCondition
   RUNG wire#powerrail
      Contact( #s10_StRecoveryCondition )
      wire#w1
      I_Contact( #sStWtResetRel )
      I_Contact( #s10_StRecoveryCondition_T1 )
      I_Contact( #s10_StRecoveryCondition_T2 )
      I_Contact( #s10_StRecoveryCondition_T3 )
      I_Contact( #s10_StRecoveryCondition_T4 )
      I_Contact( #s10_StRecoveryCondition_T5 )
      I_Contact( #s10_StRecoveryCondition_T6 )
      I_Contact( #s10_StRecoveryCondition_T7 )
      wire#w2
      Coil( #s10_StRecoveryCondition )
   END_RUNG
   RUNG wire#powerrail
      Contact( #s15_StWaitForManCorrection_T1 )
   END_RUNG wire#w1
   RUNG wire#w2
      { S7_GenerateENO := "TRUE" } Move(in := 10, out1 => #StateNo)
   END_RUNG
   // the same network as SCL:
   #s10_StRecoveryCondition := (#s10_StRecoveryCondition OR #s15_StWaitForManCorrection_T1) AND NOT #sStWtResetRel AND NOT #s10_StRecoveryCondition_T1 AND NOT #s10_StRecoveryCondition_T2 AND NOT #s10_StRecoveryCondition_T3 AND NOT #s10_StRecoveryCondition_T4 AND NOT #s10_StRecoveryCondition_T5 AND NOT #s10_StRecoveryCondition_T6 AND NOT #s10_StRecoveryCondition_T7;
   IF #s10_StRecoveryCondition THEN #StateNo := 10; END_IF;
END_REGION

REGION Network 10: Transition for STATE Num:15 StWaitForManCorrection
   RUNG wire#powerrail
      Contact( #s15_StWaitForManCorrection )
      I_Contact( #sStWtResetRel )
      Contact( #sSst )
      Contact( #iFaultReset )
      Coil( #s15_StWaitForManCorrection_T1 )
   END_RUNG
   // the same network as SCL:
   #s15_StWaitForManCorrection_T1 := #s15_StWaitForManCorrection AND NOT #sStWtResetRel AND #sSst AND #iFaultReset;
END_REGION

REGION Network 11: STATE Num:15 StWaitForManCorrection
   RUNG wire#powerrail
      Contact( #s15_StWaitForManCorrection )
      wire#w1
      I_Contact( #sStWtResetRel )
      I_Contact( #s15_StWaitForManCorrection_T1 )
      wire#w2
      Coil( #s15_StWaitForManCorrection )
   END_RUNG
   RUNG wire#powerrail
      Contact( #s10_StRecoveryCondition_T1 )
   END_RUNG wire#w1
   RUNG wire#w2
      { S7_GenerateENO := "TRUE" } Move(in := 15, out1 => #StateNo)
   END_RUNG
   // the same network as SCL:
   #s15_StWaitForManCorrection := (#s15_StWaitForManCorrection OR #s10_StRecoveryCondition_T1) AND NOT #sStWtResetRel AND NOT #s15_StWaitForManCorrection_T1;
   IF #s15_StWaitForManCorrection THEN #StateNo := 15; END_IF;
END_REGION

REGION Network 12: Transition for STATE Num:20 StChkForPalletPresent
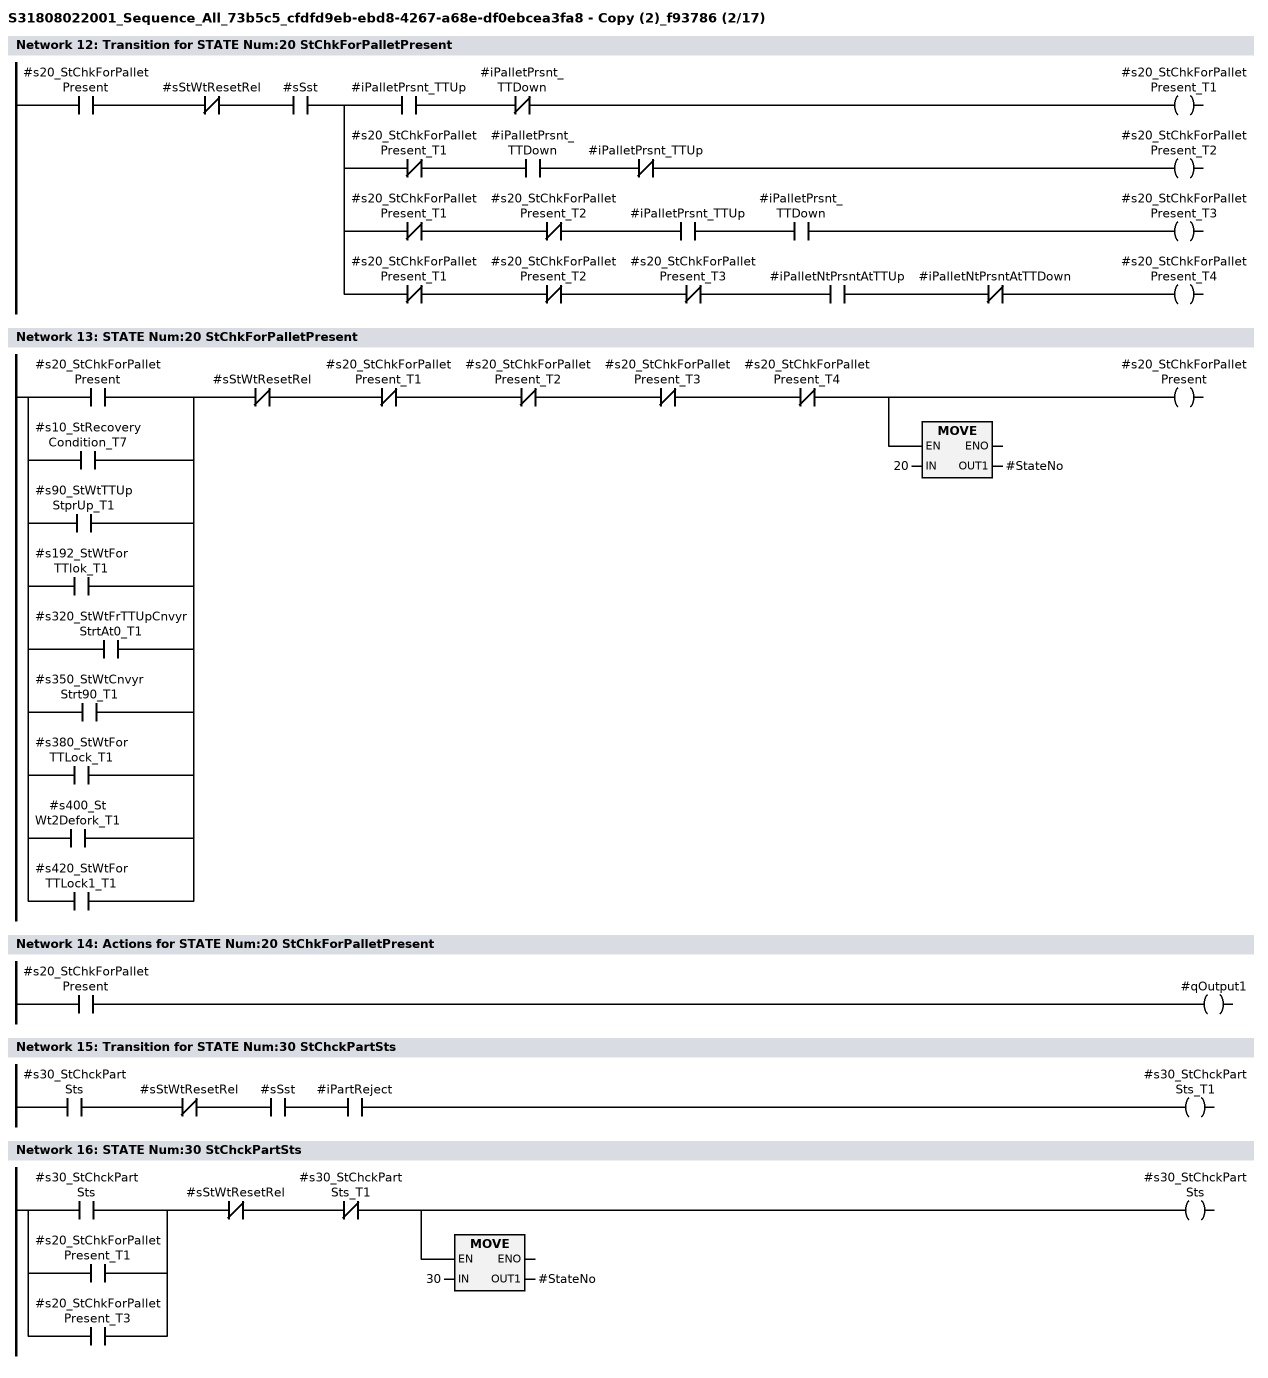
   RUNG wire#powerrail
      Contact( #s20_StChkForPalletPresent )
      I_Contact( #sStWtResetRel )
      Contact( #sSst )
      wire#w1
      Contact( #iPalletPrsnt_TTUp )
      I_Contact( #iPalletPrsnt_TTDown )
      Coil( #s20_StChkForPalletPresent_T1 )
   END_RUNG
   RUNG wire#w1
      I_Contact( #s20_StChkForPalletPresent_T1 )
      Contact( #iPalletPrsnt_TTDown )
      I_Contact( #iPalletPrsnt_TTUp )
      Coil( #s20_StChkForPalletPresent_T2 )
   END_RUNG
   RUNG wire#w1
      I_Contact( #s20_StChkForPalletPresent_T1 )
      I_Contact( #s20_StChkForPalletPresent_T2 )
      Contact( #iPalletPrsnt_TTUp )
      Contact( #iPalletPrsnt_TTDown )
      Coil( #s20_StChkForPalletPresent_T3 )
   END_RUNG
   RUNG wire#w1
      I_Contact( #s20_StChkForPalletPresent_T1 )
      I_Contact( #s20_StChkForPalletPresent_T2 )
      I_Contact( #s20_StChkForPalletPresent_T3 )
      Contact( #iPalletNtPrsntAtTTUp )
      I_Contact( #iPalletNtPrsntAtTTDown )
      Coil( #s20_StChkForPalletPresent_T4 )
   END_RUNG
   // the same network as SCL:
   #_w1 := #s20_StChkForPalletPresent AND NOT #sStWtResetRel AND #sSst;
   #s20_StChkForPalletPresent_T1 := #_w1 AND #iPalletPrsnt_TTUp AND NOT #iPalletPrsnt_TTDown;
   #s20_StChkForPalletPresent_T2 := #_w1 AND NOT #s20_StChkForPalletPresent_T1 AND #iPalletPrsnt_TTDown AND NOT #iPalletPrsnt_TTUp;
   #s20_StChkForPalletPresent_T3 := #_w1 AND NOT #s20_StChkForPalletPresent_T1 AND NOT #s20_StChkForPalletPresent_T2 AND #iPalletPrsnt_TTUp AND #iPalletPrsnt_TTDown;
   #s20_StChkForPalletPresent_T4 := #_w1 AND NOT #s20_StChkForPalletPresent_T1 AND NOT #s20_StChkForPalletPresent_T2 AND NOT #s20_StChkForPalletPresent_T3 AND #iPalletNtPrsntAtTTUp AND NOT #iPalletNtPrsntAtTTDown;
END_REGION

REGION Network 13: STATE Num:20 StChkForPalletPresent
   RUNG wire#powerrail
      Contact( #s20_StChkForPalletPresent )
      wire#w1
      I_Contact( #sStWtResetRel )
      I_Contact( #s20_StChkForPalletPresent_T1 )
      I_Contact( #s20_StChkForPalletPresent_T2 )
      I_Contact( #s20_StChkForPalletPresent_T3 )
      I_Contact( #s20_StChkForPalletPresent_T4 )
      wire#w2
      Coil( #s20_StChkForPalletPresent )
   END_RUNG
   RUNG wire#powerrail
      Contact( #s10_StRecoveryCondition_T7 )
   END_RUNG wire#w1
   RUNG wire#powerrail
      Contact( #s90_StWtTTUpStprUp_T1 )
   END_RUNG wire#w1
   RUNG wire#powerrail
      Contact( #s192_StWtForTTlok_T1 )
   END_RUNG wire#w1
   RUNG wire#powerrail
      Contact( #s320_StWtFrTTUpCnvyrStrtAt0_T1 )
   END_RUNG wire#w1
   RUNG wire#powerrail
      Contact( #s350_StWtCnvyrStrt90_T1 )
   END_RUNG wire#w1
   RUNG wire#powerrail
      Contact( #s380_StWtForTTLock_T1 )
   END_RUNG wire#w1
   RUNG wire#powerrail
      Contact( #s400_StWt2Defork_T1 )
   END_RUNG wire#w1
   RUNG wire#powerrail
      Contact( #s420_StWtForTTLock1_T1 )
   END_RUNG wire#w1
   RUNG wire#w2
      { S7_GenerateENO := "TRUE" } Move(in := 20, out1 => #StateNo)
   END_RUNG
   // the same network as SCL:
   #s20_StChkForPalletPresent := (#s20_StChkForPalletPresent OR #s10_StRecoveryCondition_T7 OR #s90_StWtTTUpStprUp_T1 OR #s192_StWtForTTlok_T1 OR #s320_StWtFrTTUpCnvyrStrtAt0_T1 OR #s350_StWtCnvyrStrt90_T1 OR #s380_StWtForTTLock_T1 OR #s400_StWt2Defork_T1 OR #s420_StWtForTTLock1_T1) AND NOT #sStWtResetRel AND NOT #s20_StChkForPalletPresent_T1 AND NOT #s20_StChkForPalletPresent_T2 AND NOT #s20_StChkForPalletPresent_T3 AND NOT #s20_StChkForPalletPresent_T4;
   IF #s20_StChkForPalletPresent THEN #StateNo := 20; END_IF;
END_REGION

REGION Network 14: Actions for STATE Num:20 StChkForPalletPresent
   RUNG wire#powerrail
      Contact( #s20_StChkForPalletPresent )
      Coil( #qOutput1 )
   END_RUNG
   // the same network as SCL:
   #qOutput1 := #s20_StChkForPalletPresent;
END_REGION

REGION Network 15: Transition for STATE Num:30 StChckPartSts
   RUNG wire#powerrail
      Contact( #s30_StChckPartSts )
      I_Contact( #sStWtResetRel )
      Contact( #sSst )
      Contact( #iPartReject )
      Coil( #s30_StChckPartSts_T1 )
   END_RUNG
   // the same network as SCL:
   #s30_StChckPartSts_T1 := #s30_StChckPartSts AND NOT #sStWtResetRel AND #sSst AND #iPartReject;
END_REGION

REGION Network 16: STATE Num:30 StChckPartSts
   RUNG wire#powerrail
      Contact( #s30_StChckPartSts )
      wire#w1
      I_Contact( #sStWtResetRel )
      I_Contact( #s30_StChckPartSts_T1 )
      wire#w2
      Coil( #s30_StChckPartSts )
   END_RUNG
   RUNG wire#powerrail
      Contact( #s20_StChkForPalletPresent_T1 )
   END_RUNG wire#w1
   RUNG wire#powerrail
      Contact( #s20_StChkForPalletPresent_T3 )
   END_RUNG wire#w1
   RUNG wire#w2
      { S7_GenerateENO := "TRUE" } Move(in := 30, out1 => #StateNo)
   END_RUNG
   // the same network as SCL:
   #s30_StChckPartSts := (#s30_StChckPartSts OR #s20_StChkForPalletPresent_T1 OR #s20_StChkForPalletPresent_T3) AND NOT #sStWtResetRel AND NOT #s30_StChckPartSts_T1;
   IF #s30_StChckPartSts THEN #StateNo := 30; END_IF;
END_REGION

REGION Network 17: Actions for STATE Num:30 StChckPartSts
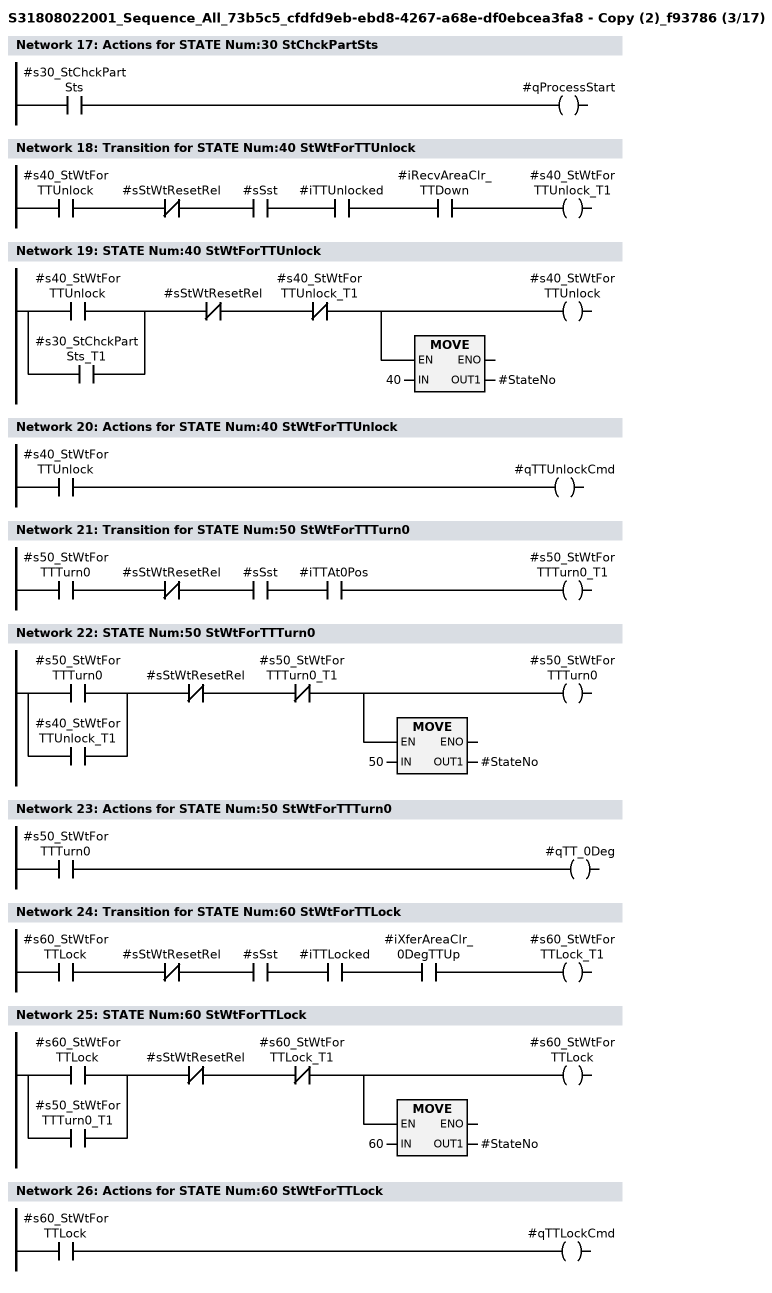
   RUNG wire#powerrail
      Contact( #s30_StChckPartSts )
      Coil( #qProcessStart )
   END_RUNG
   // the same network as SCL:
   #qProcessStart := #s30_StChckPartSts;
END_REGION

REGION Network 18: Transition for STATE Num:40 StWtForTTUnlock
   RUNG wire#powerrail
      Contact( #s40_StWtForTTUnlock )
      I_Contact( #sStWtResetRel )
      Contact( #sSst )
      Contact( #iTTUnlocked )
      Contact( #iRecvAreaClr_TTDown )
      Coil( #s40_StWtForTTUnlock_T1 )
   END_RUNG
   // the same network as SCL:
   #s40_StWtForTTUnlock_T1 := #s40_StWtForTTUnlock AND NOT #sStWtResetRel AND #sSst AND #iTTUnlocked AND #iRecvAreaClr_TTDown;
END_REGION

REGION Network 19: STATE Num:40 StWtForTTUnlock
   RUNG wire#powerrail
      Contact( #s40_StWtForTTUnlock )
      wire#w1
      I_Contact( #sStWtResetRel )
      I_Contact( #s40_StWtForTTUnlock_T1 )
      wire#w2
      Coil( #s40_StWtForTTUnlock )
   END_RUNG
   RUNG wire#powerrail
      Contact( #s30_StChckPartSts_T1 )
   END_RUNG wire#w1
   RUNG wire#w2
      { S7_GenerateENO := "TRUE" } Move(in := 40, out1 => #StateNo)
   END_RUNG
   // the same network as SCL:
   #s40_StWtForTTUnlock := (#s40_StWtForTTUnlock OR #s30_StChckPartSts_T1) AND NOT #sStWtResetRel AND NOT #s40_StWtForTTUnlock_T1;
   IF #s40_StWtForTTUnlock THEN #StateNo := 40; END_IF;
END_REGION

REGION Network 20: Actions for STATE Num:40 StWtForTTUnlock
   RUNG wire#powerrail
      Contact( #s40_StWtForTTUnlock )
      Coil( #qTTUnlockCmd )
   END_RUNG
   // the same network as SCL:
   #qTTUnlockCmd := #s40_StWtForTTUnlock;
END_REGION

REGION Network 21: Transition for STATE Num:50 StWtForTTTurn0
   RUNG wire#powerrail
      Contact( #s50_StWtForTTTurn0 )
      I_Contact( #sStWtResetRel )
      Contact( #sSst )
      Contact( #iTTAt0Pos )
      Coil( #s50_StWtForTTTurn0_T1 )
   END_RUNG
   // the same network as SCL:
   #s50_StWtForTTTurn0_T1 := #s50_StWtForTTTurn0 AND NOT #sStWtResetRel AND #sSst AND #iTTAt0Pos;
END_REGION

REGION Network 22: STATE Num:50 StWtForTTTurn0
   RUNG wire#powerrail
      Contact( #s50_StWtForTTTurn0 )
      wire#w1
      I_Contact( #sStWtResetRel )
      I_Contact( #s50_StWtForTTTurn0_T1 )
      wire#w2
      Coil( #s50_StWtForTTTurn0 )
   END_RUNG
   RUNG wire#powerrail
      Contact( #s40_StWtForTTUnlock_T1 )
   END_RUNG wire#w1
   RUNG wire#w2
      { S7_GenerateENO := "TRUE" } Move(in := 50, out1 => #StateNo)
   END_RUNG
   // the same network as SCL:
   #s50_StWtForTTTurn0 := (#s50_StWtForTTTurn0 OR #s40_StWtForTTUnlock_T1) AND NOT #sStWtResetRel AND NOT #s50_StWtForTTTurn0_T1;
   IF #s50_StWtForTTTurn0 THEN #StateNo := 50; END_IF;
END_REGION

REGION Network 23: Actions for STATE Num:50 StWtForTTTurn0
   RUNG wire#powerrail
      Contact( #s50_StWtForTTTurn0 )
      Coil( #qTT_0Deg )
   END_RUNG
   // the same network as SCL:
   #qTT_0Deg := #s50_StWtForTTTurn0;
END_REGION

REGION Network 24: Transition for STATE Num:60 StWtForTTLock
   RUNG wire#powerrail
      Contact( #s60_StWtForTTLock )
      I_Contact( #sStWtResetRel )
      Contact( #sSst )
      Contact( #iTTLocked )
      Contact( #iXferAreaClr_0DegTTUp )
      Coil( #s60_StWtForTTLock_T1 )
   END_RUNG
   // the same network as SCL:
   #s60_StWtForTTLock_T1 := #s60_StWtForTTLock AND NOT #sStWtResetRel AND #sSst AND #iTTLocked AND #iXferAreaClr_0DegTTUp;
END_REGION

REGION Network 25: STATE Num:60 StWtForTTLock
   RUNG wire#powerrail
      Contact( #s60_StWtForTTLock )
      wire#w1
      I_Contact( #sStWtResetRel )
      I_Contact( #s60_StWtForTTLock_T1 )
      wire#w2
      Coil( #s60_StWtForTTLock )
   END_RUNG
   RUNG wire#powerrail
      Contact( #s50_StWtForTTTurn0_T1 )
   END_RUNG wire#w1
   RUNG wire#w2
      { S7_GenerateENO := "TRUE" } Move(in := 60, out1 => #StateNo)
   END_RUNG
   // the same network as SCL:
   #s60_StWtForTTLock := (#s60_StWtForTTLock OR #s50_StWtForTTTurn0_T1) AND NOT #sStWtResetRel AND NOT #s60_StWtForTTLock_T1;
   IF #s60_StWtForTTLock THEN #StateNo := 60; END_IF;
END_REGION

REGION Network 26: Actions for STATE Num:60 StWtForTTLock
   RUNG wire#powerrail
      Contact( #s60_StWtForTTLock )
      Coil( #qTTLockCmd )
   END_RUNG
   // the same network as SCL:
   #qTTLockCmd := #s60_StWtForTTLock;
END_REGION

REGION Network 27: Transition for STATE Num:70 StWtOTSfrmTTUp
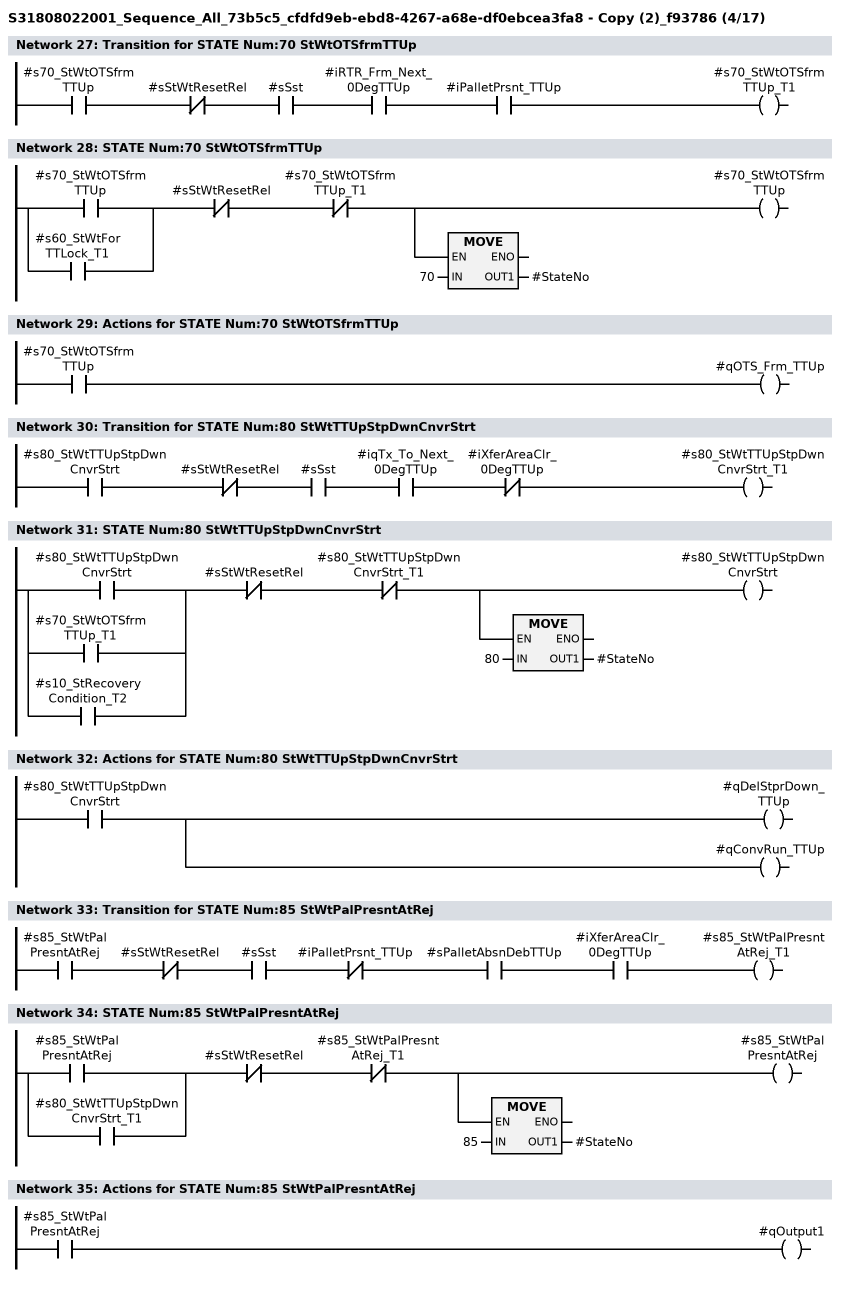
   RUNG wire#powerrail
      Contact( #s70_StWtOTSfrmTTUp )
      I_Contact( #sStWtResetRel )
      Contact( #sSst )
      Contact( #iRTR_Frm_Next_0DegTTUp )
      Contact( #iPalletPrsnt_TTUp )
      Coil( #s70_StWtOTSfrmTTUp_T1 )
   END_RUNG
   // the same network as SCL:
   #s70_StWtOTSfrmTTUp_T1 := #s70_StWtOTSfrmTTUp AND NOT #sStWtResetRel AND #sSst AND #iRTR_Frm_Next_0DegTTUp AND #iPalletPrsnt_TTUp;
END_REGION

REGION Network 28: STATE Num:70 StWtOTSfrmTTUp
   RUNG wire#powerrail
      Contact( #s70_StWtOTSfrmTTUp )
      wire#w1
      I_Contact( #sStWtResetRel )
      I_Contact( #s70_StWtOTSfrmTTUp_T1 )
      wire#w2
      Coil( #s70_StWtOTSfrmTTUp )
   END_RUNG
   RUNG wire#powerrail
      Contact( #s60_StWtForTTLock_T1 )
   END_RUNG wire#w1
   RUNG wire#w2
      { S7_GenerateENO := "TRUE" } Move(in := 70, out1 => #StateNo)
   END_RUNG
   // the same network as SCL:
   #s70_StWtOTSfrmTTUp := (#s70_StWtOTSfrmTTUp OR #s60_StWtForTTLock_T1) AND NOT #sStWtResetRel AND NOT #s70_StWtOTSfrmTTUp_T1;
   IF #s70_StWtOTSfrmTTUp THEN #StateNo := 70; END_IF;
END_REGION

REGION Network 29: Actions for STATE Num:70 StWtOTSfrmTTUp
   RUNG wire#powerrail
      Contact( #s70_StWtOTSfrmTTUp )
      Coil( #qOTS_Frm_TTUp )
   END_RUNG
   // the same network as SCL:
   #qOTS_Frm_TTUp := #s70_StWtOTSfrmTTUp;
END_REGION

REGION Network 30: Transition for STATE Num:80 StWtTTUpStpDwnCnvrStrt
   RUNG wire#powerrail
      Contact( #s80_StWtTTUpStpDwnCnvrStrt )
      I_Contact( #sStWtResetRel )
      Contact( #sSst )
      Contact( #iqTx_To_Next_0DegTTUp )
      I_Contact( #iXferAreaClr_0DegTTUp )
      Coil( #s80_StWtTTUpStpDwnCnvrStrt_T1 )
   END_RUNG
   // the same network as SCL:
   #s80_StWtTTUpStpDwnCnvrStrt_T1 := #s80_StWtTTUpStpDwnCnvrStrt AND NOT #sStWtResetRel AND #sSst AND #iqTx_To_Next_0DegTTUp AND NOT #iXferAreaClr_0DegTTUp;
END_REGION

REGION Network 31: STATE Num:80 StWtTTUpStpDwnCnvrStrt
   RUNG wire#powerrail
      Contact( #s80_StWtTTUpStpDwnCnvrStrt )
      wire#w1
      I_Contact( #sStWtResetRel )
      I_Contact( #s80_StWtTTUpStpDwnCnvrStrt_T1 )
      wire#w2
      Coil( #s80_StWtTTUpStpDwnCnvrStrt )
   END_RUNG
   RUNG wire#powerrail
      Contact( #s70_StWtOTSfrmTTUp_T1 )
   END_RUNG wire#w1
   RUNG wire#powerrail
      Contact( #s10_StRecoveryCondition_T2 )
   END_RUNG wire#w1
   RUNG wire#w2
      { S7_GenerateENO := "TRUE" } Move(in := 80, out1 => #StateNo)
   END_RUNG
   // the same network as SCL:
   #s80_StWtTTUpStpDwnCnvrStrt := (#s80_StWtTTUpStpDwnCnvrStrt OR #s70_StWtOTSfrmTTUp_T1 OR #s10_StRecoveryCondition_T2) AND NOT #sStWtResetRel AND NOT #s80_StWtTTUpStpDwnCnvrStrt_T1;
   IF #s80_StWtTTUpStpDwnCnvrStrt THEN #StateNo := 80; END_IF;
END_REGION

REGION Network 32: Actions for STATE Num:80 StWtTTUpStpDwnCnvrStrt
   RUNG wire#powerrail
      Contact( #s80_StWtTTUpStpDwnCnvrStrt )
      wire#w1
      Coil( #qDelStprDown_TTUp )
   END_RUNG
   RUNG wire#w1
      Coil( #qConvRun_TTUp )
   END_RUNG
   // the same network as SCL:
   #qDelStprDown_TTUp := #s80_StWtTTUpStpDwnCnvrStrt;
   #qConvRun_TTUp := #s80_StWtTTUpStpDwnCnvrStrt;
END_REGION

REGION Network 33: Transition for STATE Num:85 StWtPalPresntAtRej
   RUNG wire#powerrail
      Contact( #s85_StWtPalPresntAtRej )
      I_Contact( #sStWtResetRel )
      Contact( #sSst )
      I_Contact( #iPalletPrsnt_TTUp )
      Contact( #sPalletAbsnDebTTUp )
      Contact( #iXferAreaClr_0DegTTUp )
      Coil( #s85_StWtPalPresntAtRej_T1 )
   END_RUNG
   // the same network as SCL:
   #s85_StWtPalPresntAtRej_T1 := #s85_StWtPalPresntAtRej AND NOT #sStWtResetRel AND #sSst AND NOT #iPalletPrsnt_TTUp AND #sPalletAbsnDebTTUp AND #iXferAreaClr_0DegTTUp;
END_REGION

REGION Network 34: STATE Num:85 StWtPalPresntAtRej
   RUNG wire#powerrail
      Contact( #s85_StWtPalPresntAtRej )
      wire#w1
      I_Contact( #sStWtResetRel )
      I_Contact( #s85_StWtPalPresntAtRej_T1 )
      wire#w2
      Coil( #s85_StWtPalPresntAtRej )
   END_RUNG
   RUNG wire#powerrail
      Contact( #s80_StWtTTUpStpDwnCnvrStrt_T1 )
   END_RUNG wire#w1
   RUNG wire#w2
      { S7_GenerateENO := "TRUE" } Move(in := 85, out1 => #StateNo)
   END_RUNG
   // the same network as SCL:
   #s85_StWtPalPresntAtRej := (#s85_StWtPalPresntAtRej OR #s80_StWtTTUpStpDwnCnvrStrt_T1) AND NOT #sStWtResetRel AND NOT #s85_StWtPalPresntAtRej_T1;
   IF #s85_StWtPalPresntAtRej THEN #StateNo := 85; END_IF;
END_REGION

REGION Network 35: Actions for STATE Num:85 StWtPalPresntAtRej
   RUNG wire#powerrail
      Contact( #s85_StWtPalPresntAtRej )
      Coil( #qOutput1 )
   END_RUNG
   // the same network as SCL:
   #qOutput1 := #s85_StWtPalPresntAtRej;
END_REGION

REGION Network 36: Transition for STATE Num:90 StWtTTUpStprUp
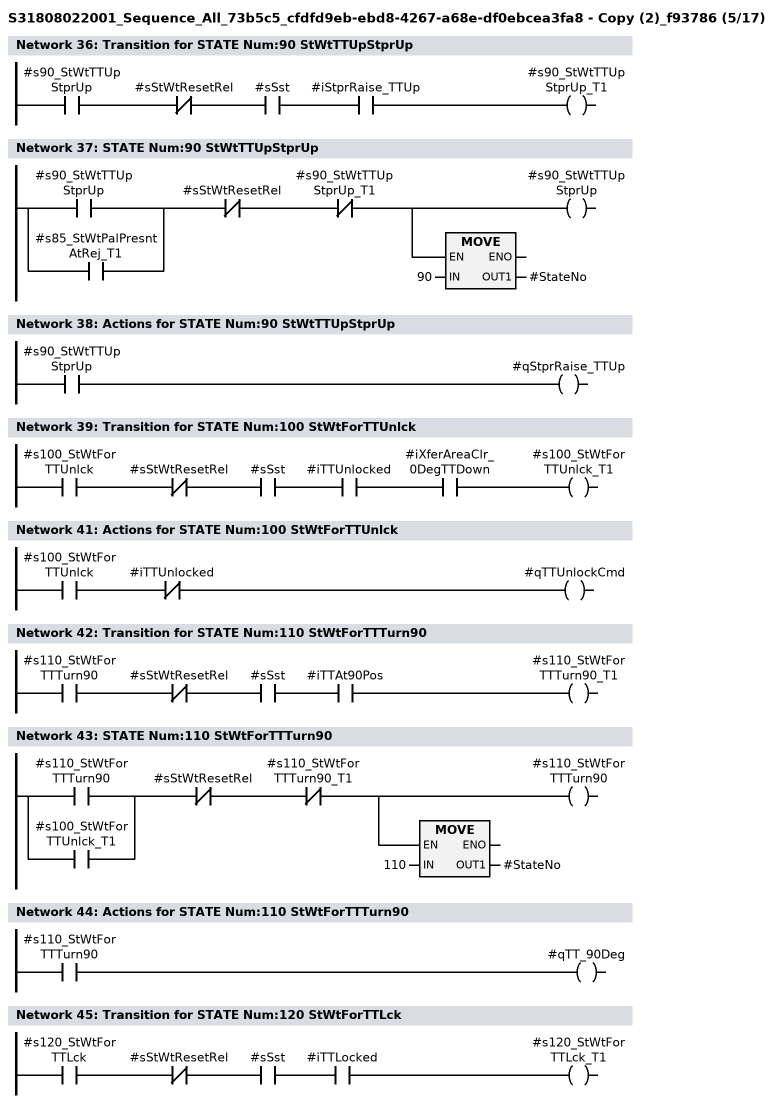
   RUNG wire#powerrail
      Contact( #s90_StWtTTUpStprUp )
      I_Contact( #sStWtResetRel )
      Contact( #sSst )
      Contact( #iStprRaise_TTUp )
      Coil( #s90_StWtTTUpStprUp_T1 )
   END_RUNG
   // the same network as SCL:
   #s90_StWtTTUpStprUp_T1 := #s90_StWtTTUpStprUp AND NOT #sStWtResetRel AND #sSst AND #iStprRaise_TTUp;
END_REGION

REGION Network 37: STATE Num:90 StWtTTUpStprUp
   RUNG wire#powerrail
      Contact( #s90_StWtTTUpStprUp )
      wire#w1
      I_Contact( #sStWtResetRel )
      I_Contact( #s90_StWtTTUpStprUp_T1 )
      wire#w2
      Coil( #s90_StWtTTUpStprUp )
   END_RUNG
   RUNG wire#powerrail
      Contact( #s85_StWtPalPresntAtRej_T1 )
   END_RUNG wire#w1
   RUNG wire#w2
      { S7_GenerateENO := "TRUE" } Move(in := 90, out1 => #StateNo)
   END_RUNG
   // the same network as SCL:
   #s90_StWtTTUpStprUp := (#s90_StWtTTUpStprUp OR #s85_StWtPalPresntAtRej_T1) AND NOT #sStWtResetRel AND NOT #s90_StWtTTUpStprUp_T1;
   IF #s90_StWtTTUpStprUp THEN #StateNo := 90; END_IF;
END_REGION

REGION Network 38: Actions for STATE Num:90 StWtTTUpStprUp
   RUNG wire#powerrail
      Contact( #s90_StWtTTUpStprUp )
      Coil( #qStprRaise_TTUp )
   END_RUNG
   // the same network as SCL:
   #qStprRaise_TTUp := #s90_StWtTTUpStprUp;
END_REGION

REGION Network 39: Transition for STATE Num:100 StWtForTTUnlck
   RUNG wire#powerrail
      Contact( #s100_StWtForTTUnlck )
      I_Contact( #sStWtResetRel )
      Contact( #sSst )
      Contact( #iTTUnlocked )
      Contact( #iXferAreaClr_0DegTTDown )
      Coil( #s100_StWtForTTUnlck_T1 )
   END_RUNG
   // the same network as SCL:
   #s100_StWtForTTUnlck_T1 := #s100_StWtForTTUnlck AND NOT #sStWtResetRel AND #sSst AND #iTTUnlocked AND #iXferAreaClr_0DegTTDown;
END_REGION

REGION Network 40 (STL): STATE Num:100 StWtForTTUnlck
         A(;
         O     #s100_StWtForTTUnlck;
         );
         AN    #sStWtResetRel;
         AN    #s100_StWtForTTUnlck_T1;
         =     <??.?>;
         A     <??.?>;
         BLD   102;
         =     #s100_StWtForTTUnlck;
         A     <??.?>;
         JNB   Label_13;
         L     100;
         T     #StateNo;
   Label_13:NOP   0;
END_REGION

REGION Network 41: Actions for STATE Num:100 StWtForTTUnlck
   RUNG wire#powerrail
      Contact( #s100_StWtForTTUnlck )
      I_Contact( #iTTUnlocked )
      Coil( #qTTUnlockCmd )
   END_RUNG
   // the same network as SCL:
   #qTTUnlockCmd := #s100_StWtForTTUnlck AND NOT #iTTUnlocked;
END_REGION

REGION Network 42: Transition for STATE Num:110 StWtForTTTurn90
   RUNG wire#powerrail
      Contact( #s110_StWtForTTTurn90 )
      I_Contact( #sStWtResetRel )
      Contact( #sSst )
      Contact( #iTTAt90Pos )
      Coil( #s110_StWtForTTTurn90_T1 )
   END_RUNG
   // the same network as SCL:
   #s110_StWtForTTTurn90_T1 := #s110_StWtForTTTurn90 AND NOT #sStWtResetRel AND #sSst AND #iTTAt90Pos;
END_REGION

REGION Network 43: STATE Num:110 StWtForTTTurn90
   RUNG wire#powerrail
      Contact( #s110_StWtForTTTurn90 )
      wire#w1
      I_Contact( #sStWtResetRel )
      I_Contact( #s110_StWtForTTTurn90_T1 )
      wire#w2
      Coil( #s110_StWtForTTTurn90 )
   END_RUNG
   RUNG wire#powerrail
      Contact( #s100_StWtForTTUnlck_T1 )
   END_RUNG wire#w1
   RUNG wire#w2
      { S7_GenerateENO := "TRUE" } Move(in := 110, out1 => #StateNo)
   END_RUNG
   // the same network as SCL:
   #s110_StWtForTTTurn90 := (#s110_StWtForTTTurn90 OR #s100_StWtForTTUnlck_T1) AND NOT #sStWtResetRel AND NOT #s110_StWtForTTTurn90_T1;
   IF #s110_StWtForTTTurn90 THEN #StateNo := 110; END_IF;
END_REGION

REGION Network 44: Actions for STATE Num:110 StWtForTTTurn90
   RUNG wire#powerrail
      Contact( #s110_StWtForTTTurn90 )
      Coil( #qTT_90Deg )
   END_RUNG
   // the same network as SCL:
   #qTT_90Deg := #s110_StWtForTTTurn90;
END_REGION

REGION Network 45: Transition for STATE Num:120 StWtForTTLck
   RUNG wire#powerrail
      Contact( #s120_StWtForTTLck )
      I_Contact( #sStWtResetRel )
      Contact( #sSst )
      Contact( #iTTLocked )
      Coil( #s120_StWtForTTLck_T1 )
   END_RUNG
   // the same network as SCL:
   #s120_StWtForTTLck_T1 := #s120_StWtForTTLck AND NOT #sStWtResetRel AND #sSst AND #iTTLocked;
END_REGION

REGION Network 46: STATE Num:120 StWtForTTLck
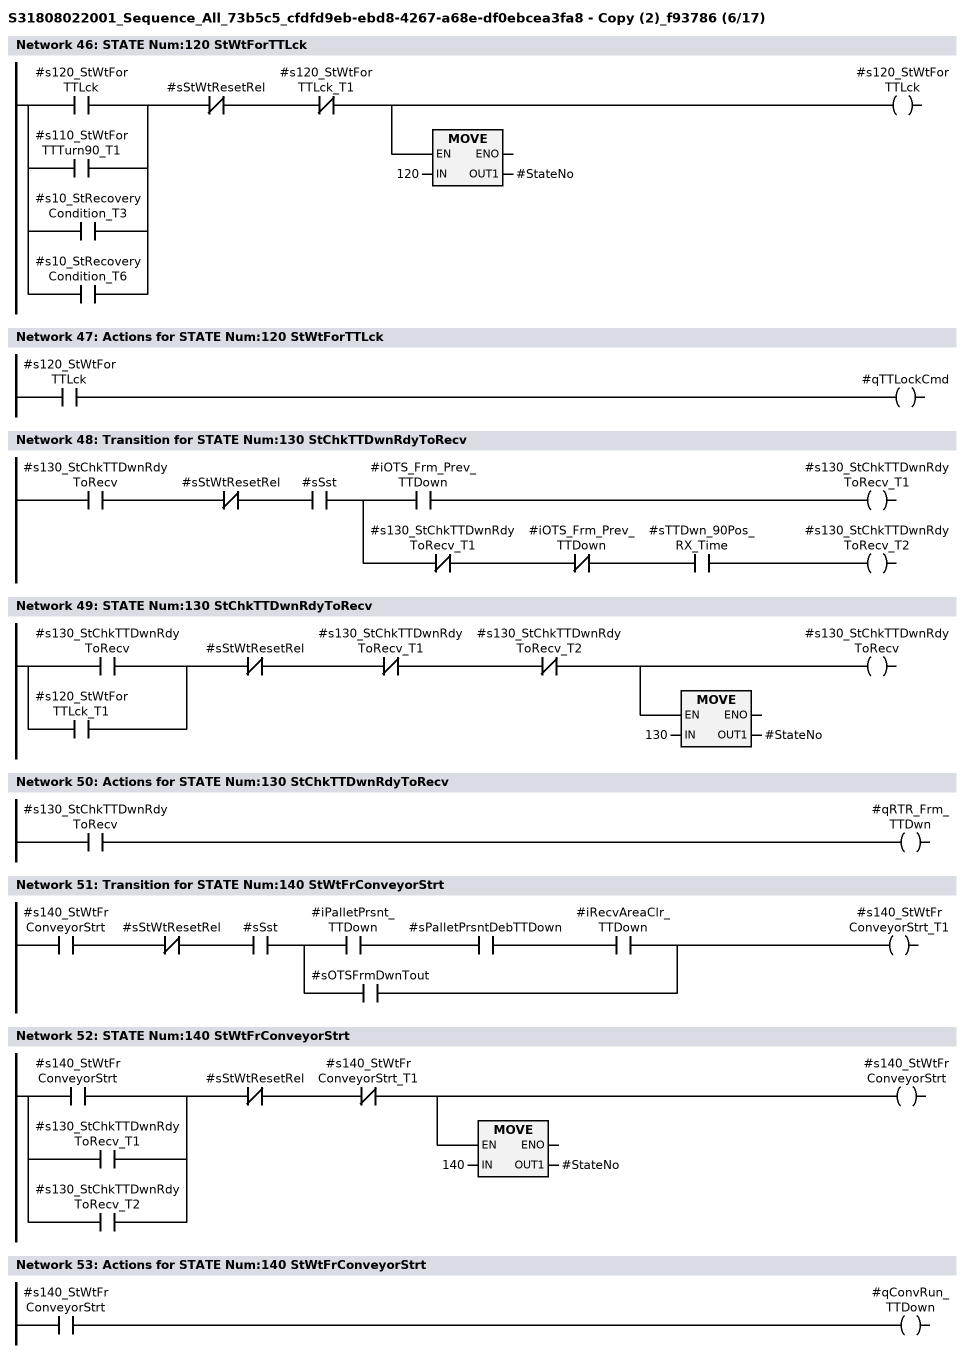
   RUNG wire#powerrail
      Contact( #s120_StWtForTTLck )
      wire#w1
      I_Contact( #sStWtResetRel )
      I_Contact( #s120_StWtForTTLck_T1 )
      wire#w2
      Coil( #s120_StWtForTTLck )
   END_RUNG
   RUNG wire#powerrail
      Contact( #s110_StWtForTTTurn90_T1 )
   END_RUNG wire#w1
   RUNG wire#powerrail
      Contact( #s10_StRecoveryCondition_T3 )
   END_RUNG wire#w1
   RUNG wire#powerrail
      Contact( #s10_StRecoveryCondition_T6 )
   END_RUNG wire#w1
   RUNG wire#w2
      { S7_GenerateENO := "TRUE" } Move(in := 120, out1 => #StateNo)
   END_RUNG
   // the same network as SCL:
   #s120_StWtForTTLck := (#s120_StWtForTTLck OR #s110_StWtForTTTurn90_T1 OR #s10_StRecoveryCondition_T3 OR #s10_StRecoveryCondition_T6) AND NOT #sStWtResetRel AND NOT #s120_StWtForTTLck_T1;
   IF #s120_StWtForTTLck THEN #StateNo := 120; END_IF;
END_REGION

REGION Network 47: Actions for STATE Num:120 StWtForTTLck
   RUNG wire#powerrail
      Contact( #s120_StWtForTTLck )
      Coil( #qTTLockCmd )
   END_RUNG
   // the same network as SCL:
   #qTTLockCmd := #s120_StWtForTTLck;
END_REGION

REGION Network 48: Transition for STATE Num:130 StChkTTDwnRdyToRecv
   RUNG wire#powerrail
      Contact( #s130_StChkTTDwnRdyToRecv )
      I_Contact( #sStWtResetRel )
      Contact( #sSst )
      wire#w1
      Contact( #iOTS_Frm_Prev_TTDown )
      Coil( #s130_StChkTTDwnRdyToRecv_T1 )
   END_RUNG
   RUNG wire#w1
      I_Contact( #s130_StChkTTDwnRdyToRecv_T1 )
      I_Contact( #iOTS_Frm_Prev_TTDown )
      Contact( #sTTDwn_90Pos_RX_Time )
      Coil( #s130_StChkTTDwnRdyToRecv_T2 )
   END_RUNG
   // the same network as SCL:
   #_w1 := #s130_StChkTTDwnRdyToRecv AND NOT #sStWtResetRel AND #sSst;
   #s130_StChkTTDwnRdyToRecv_T1 := #_w1 AND #iOTS_Frm_Prev_TTDown;
   #s130_StChkTTDwnRdyToRecv_T2 := #_w1 AND NOT #s130_StChkTTDwnRdyToRecv_T1 AND NOT #iOTS_Frm_Prev_TTDown AND #sTTDwn_90Pos_RX_Time;
END_REGION

REGION Network 49: STATE Num:130 StChkTTDwnRdyToRecv
   RUNG wire#powerrail
      Contact( #s130_StChkTTDwnRdyToRecv )
      wire#w1
      I_Contact( #sStWtResetRel )
      I_Contact( #s130_StChkTTDwnRdyToRecv_T1 )
      I_Contact( #s130_StChkTTDwnRdyToRecv_T2 )
      wire#w2
      Coil( #s130_StChkTTDwnRdyToRecv )
   END_RUNG
   RUNG wire#powerrail
      Contact( #s120_StWtForTTLck_T1 )
   END_RUNG wire#w1
   RUNG wire#w2
      { S7_GenerateENO := "TRUE" } Move(in := 130, out1 => #StateNo)
   END_RUNG
   // the same network as SCL:
   #s130_StChkTTDwnRdyToRecv := (#s130_StChkTTDwnRdyToRecv OR #s120_StWtForTTLck_T1) AND NOT #sStWtResetRel AND NOT #s130_StChkTTDwnRdyToRecv_T1 AND NOT #s130_StChkTTDwnRdyToRecv_T2;
   IF #s130_StChkTTDwnRdyToRecv THEN #StateNo := 130; END_IF;
END_REGION

REGION Network 50: Actions for STATE Num:130 StChkTTDwnRdyToRecv
   RUNG wire#powerrail
      Contact( #s130_StChkTTDwnRdyToRecv )
      Coil( #qRTR_Frm_TTDwn )
   END_RUNG
   // the same network as SCL:
   #qRTR_Frm_TTDwn := #s130_StChkTTDwnRdyToRecv;
END_REGION

REGION Network 51: Transition for STATE Num:140 StWtFrConveyorStrt
   RUNG wire#powerrail
      Contact( #s140_StWtFrConveyorStrt )
      I_Contact( #sStWtResetRel )
      Contact( #sSst )
      wire#w1
      Contact( #iPalletPrsnt_TTDown )
      Contact( #sPalletPrsntDebTTDown )
      Contact( #iRecvAreaClr_TTDown )
      wire#w2
      Coil( #s140_StWtFrConveyorStrt_T1 )
   END_RUNG
   RUNG wire#w1
      Contact( #sOTSFrmDwnTout )
   END_RUNG wire#w2
   // the same network as SCL:
   #s140_StWtFrConveyorStrt_T1 := #s140_StWtFrConveyorStrt AND NOT #sStWtResetRel AND #sSst AND ((#iPalletPrsnt_TTDown AND #sPalletPrsntDebTTDown AND #iRecvAreaClr_TTDown) OR #sOTSFrmDwnTout);
END_REGION

REGION Network 52: STATE Num:140 StWtFrConveyorStrt
   RUNG wire#powerrail
      Contact( #s140_StWtFrConveyorStrt )
      wire#w1
      I_Contact( #sStWtResetRel )
      I_Contact( #s140_StWtFrConveyorStrt_T1 )
      wire#w2
      Coil( #s140_StWtFrConveyorStrt )
   END_RUNG
   RUNG wire#powerrail
      Contact( #s130_StChkTTDwnRdyToRecv_T1 )
   END_RUNG wire#w1
   RUNG wire#powerrail
      Contact( #s130_StChkTTDwnRdyToRecv_T2 )
   END_RUNG wire#w1
   RUNG wire#w2
      { S7_GenerateENO := "TRUE" } Move(in := 140, out1 => #StateNo)
   END_RUNG
   // the same network as SCL:
   #s140_StWtFrConveyorStrt := (#s140_StWtFrConveyorStrt OR #s130_StChkTTDwnRdyToRecv_T1 OR #s130_StChkTTDwnRdyToRecv_T2) AND NOT #sStWtResetRel AND NOT #s140_StWtFrConveyorStrt_T1;
   IF #s140_StWtFrConveyorStrt THEN #StateNo := 140; END_IF;
END_REGION

REGION Network 53: Actions for STATE Num:140 StWtFrConveyorStrt
   RUNG wire#powerrail
      Contact( #s140_StWtFrConveyorStrt )
      Coil( #qConvRun_TTDown )
   END_RUNG
   // the same network as SCL:
   #qConvRun_TTDown := #s140_StWtFrConveyorStrt;
END_REGION

REGION Network 54: Transition for STATE Num:150 StChkNxtStRdyToRecvTTUp
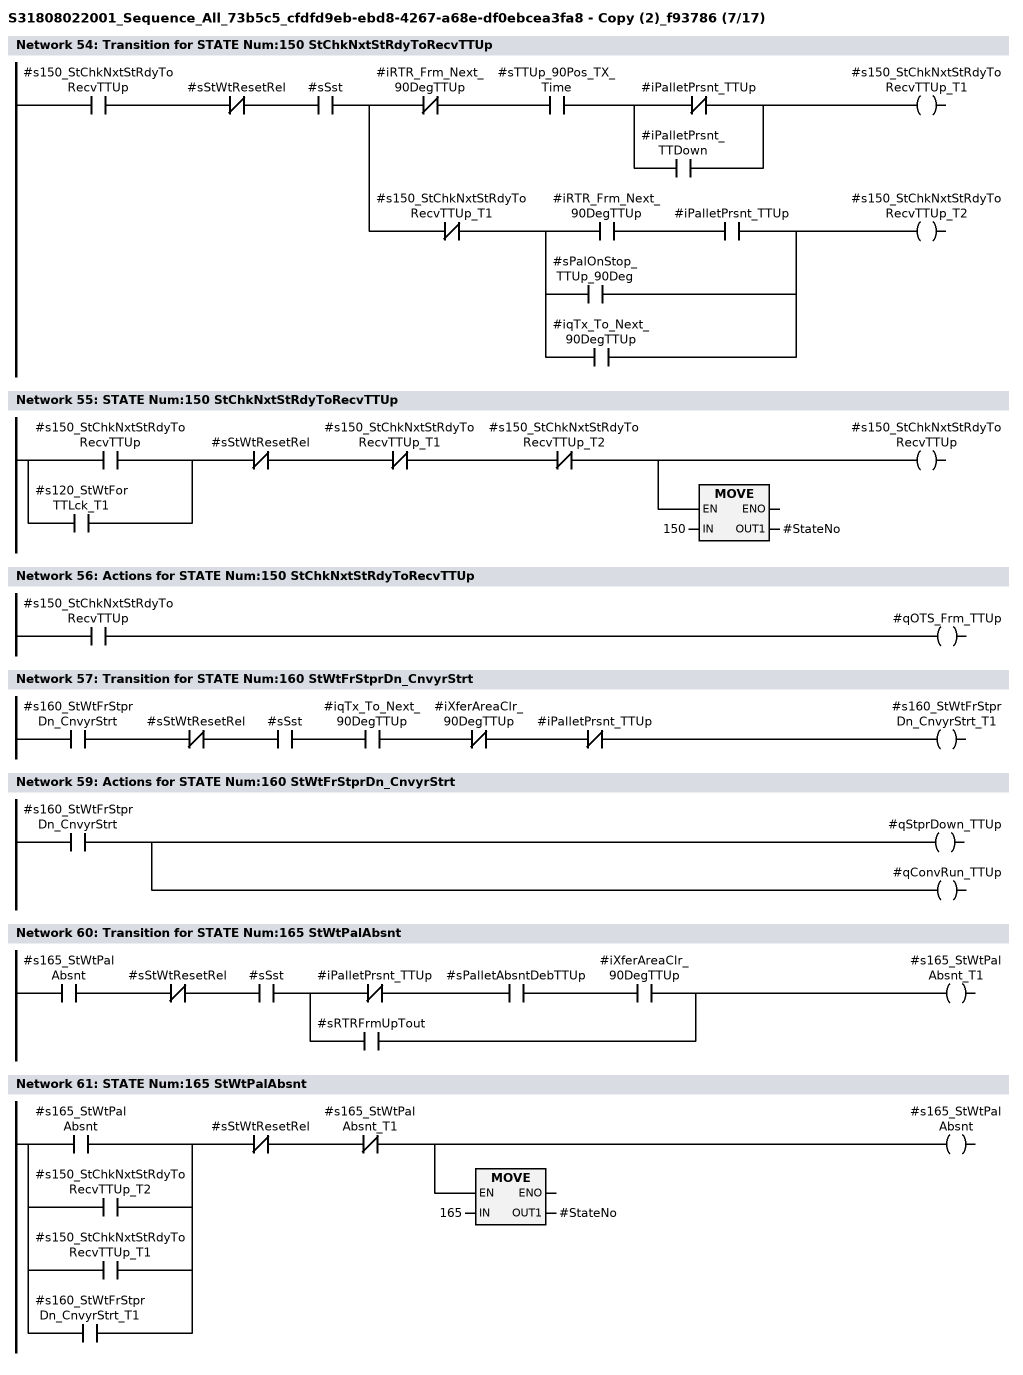
   RUNG wire#powerrail
      Contact( #s150_StChkNxtStRdyToRecvTTUp )
      I_Contact( #sStWtResetRel )
      Contact( #sSst )
      wire#w1
      I_Contact( #iRTR_Frm_Next_90DegTTUp )
      Contact( #sTTUp_90Pos_TX_Time )
      wire#w2
      I_Contact( #iPalletPrsnt_TTUp )
      wire#w3
      Coil( #s150_StChkNxtStRdyToRecvTTUp_T1 )
   END_RUNG
   RUNG wire#w2
      Contact( #iPalletPrsnt_TTDown )
   END_RUNG wire#w3
   RUNG wire#w1
      I_Contact( #s150_StChkNxtStRdyToRecvTTUp_T1 )
      wire#w4
      Contact( #iRTR_Frm_Next_90DegTTUp )
      Contact( #iPalletPrsnt_TTUp )
      wire#w5
      Coil( #s150_StChkNxtStRdyToRecvTTUp_T2 )
   END_RUNG
   RUNG wire#w4
      Contact( #sPalOnStop_TTUp_90Deg )
   END_RUNG wire#w5
   RUNG wire#w4
      Contact( #iqTx_To_Next_90DegTTUp )
   END_RUNG wire#w5
   // the same network as SCL:
   #_w1 := #s150_StChkNxtStRdyToRecvTTUp AND NOT #sStWtResetRel AND #sSst;
   #s150_StChkNxtStRdyToRecvTTUp_T1 := #_w1 AND NOT #iRTR_Frm_Next_90DegTTUp AND #sTTUp_90Pos_TX_Time AND (NOT #iPalletPrsnt_TTUp OR #iPalletPrsnt_TTDown);
   #s150_StChkNxtStRdyToRecvTTUp_T2 := #_w1 AND NOT #s150_StChkNxtStRdyToRecvTTUp_T1 AND ((#iRTR_Frm_Next_90DegTTUp AND #iPalletPrsnt_TTUp) OR #sPalOnStop_TTUp_90Deg OR #iqTx_To_Next_90DegTTUp);
END_REGION

REGION Network 55: STATE Num:150 StChkNxtStRdyToRecvTTUp
   RUNG wire#powerrail
      Contact( #s150_StChkNxtStRdyToRecvTTUp )
      wire#w1
      I_Contact( #sStWtResetRel )
      I_Contact( #s150_StChkNxtStRdyToRecvTTUp_T1 )
      I_Contact( #s150_StChkNxtStRdyToRecvTTUp_T2 )
      wire#w2
      Coil( #s150_StChkNxtStRdyToRecvTTUp )
   END_RUNG
   RUNG wire#powerrail
      Contact( #s120_StWtForTTLck_T1 )
   END_RUNG wire#w1
   RUNG wire#w2
      { S7_GenerateENO := "TRUE" } Move(in := 150, out1 => #StateNo)
   END_RUNG
   // the same network as SCL:
   #s150_StChkNxtStRdyToRecvTTUp := (#s150_StChkNxtStRdyToRecvTTUp OR #s120_StWtForTTLck_T1) AND NOT #sStWtResetRel AND NOT #s150_StChkNxtStRdyToRecvTTUp_T1 AND NOT #s150_StChkNxtStRdyToRecvTTUp_T2;
   IF #s150_StChkNxtStRdyToRecvTTUp THEN #StateNo := 150; END_IF;
END_REGION

REGION Network 56: Actions for STATE Num:150 StChkNxtStRdyToRecvTTUp
   RUNG wire#powerrail
      Contact( #s150_StChkNxtStRdyToRecvTTUp )
      Coil( #qOTS_Frm_TTUp )
   END_RUNG
   // the same network as SCL:
   #qOTS_Frm_TTUp := #s150_StChkNxtStRdyToRecvTTUp;
END_REGION

REGION Network 57: Transition for STATE Num:160 StWtFrStprDn_CnvyrStrt
   RUNG wire#powerrail
      Contact( #s160_StWtFrStprDn_CnvyrStrt )
      I_Contact( #sStWtResetRel )
      Contact( #sSst )
      Contact( #iqTx_To_Next_90DegTTUp )
      I_Contact( #iXferAreaClr_90DegTTUp )
      I_Contact( #iPalletPrsnt_TTUp )
      Coil( #s160_StWtFrStprDn_CnvyrStrt_T1 )
   END_RUNG
   // the same network as SCL:
   #s160_StWtFrStprDn_CnvyrStrt_T1 := #s160_StWtFrStprDn_CnvyrStrt AND NOT #sStWtResetRel AND #sSst AND #iqTx_To_Next_90DegTTUp AND NOT #iXferAreaClr_90DegTTUp AND NOT #iPalletPrsnt_TTUp;
END_REGION

REGION Network 58 (STL): STATE Num:160 StWtFrStprDn_CnvyrStrt
         A(;
         O     #s160_StWtFrStprDn_CnvyrStrt;
   //wrong transition variable removed
         );
         AN    #sStWtResetRel;
         AN    #s160_StWtFrStprDn_CnvyrStrt_T1;
         =     <??.?>;
         A     <??.?>;
         BLD   102;
         =     #s160_StWtFrStprDn_CnvyrStrt;
         A     <??.?>;
         JNB   Label_19;
         L     160;
         T     #StateNo;
   Label_19:NOP   0;
END_REGION

REGION Network 59: Actions for STATE Num:160 StWtFrStprDn_CnvyrStrt
   RUNG wire#powerrail
      Contact( #s160_StWtFrStprDn_CnvyrStrt )
      wire#w1
      Coil( #qStprDown_TTUp )
   END_RUNG
   RUNG wire#w1
      Coil( #qConvRun_TTUp )
   END_RUNG
   // the same network as SCL:
   #qStprDown_TTUp := #s160_StWtFrStprDn_CnvyrStrt;
   #qConvRun_TTUp := #s160_StWtFrStprDn_CnvyrStrt;
END_REGION

REGION Network 60: Transition for STATE Num:165 StWtPalAbsnt
   RUNG wire#powerrail
      Contact( #s165_StWtPalAbsnt )
      I_Contact( #sStWtResetRel )
      Contact( #sSst )
      wire#w1
      I_Contact( #iPalletPrsnt_TTUp )
      Contact( #sPalletAbsntDebTTUp )
      Contact( #iXferAreaClr_90DegTTUp )
      wire#w2
      Coil( #s165_StWtPalAbsnt_T1 )
   END_RUNG
   RUNG wire#w1
      Contact( #sRTRFrmUpTout )
   END_RUNG wire#w2
   // the same network as SCL:
   #s165_StWtPalAbsnt_T1 := #s165_StWtPalAbsnt AND NOT #sStWtResetRel AND #sSst AND ((NOT #iPalletPrsnt_TTUp AND #sPalletAbsntDebTTUp AND #iXferAreaClr_90DegTTUp) OR #sRTRFrmUpTout);
END_REGION

REGION Network 61: STATE Num:165 StWtPalAbsnt
   RUNG wire#powerrail
      Contact( #s165_StWtPalAbsnt )
      wire#w1
      I_Contact( #sStWtResetRel )
      I_Contact( #s165_StWtPalAbsnt_T1 )
      wire#w2
      Coil( #s165_StWtPalAbsnt )
   END_RUNG
   RUNG wire#powerrail
      Contact( #s150_StChkNxtStRdyToRecvTTUp_T2 )
   END_RUNG wire#w1
   RUNG wire#powerrail
      Contact( #s150_StChkNxtStRdyToRecvTTUp_T1 )
   END_RUNG wire#w1
   RUNG wire#powerrail
      Contact( #s160_StWtFrStprDn_CnvyrStrt_T1 )
   END_RUNG wire#w1
   RUNG wire#w2
      { S7_GenerateENO := "TRUE" } Move(in := 165, out1 => #StateNo)
   END_RUNG
   // the same network as SCL:
   #s165_StWtPalAbsnt := (#s165_StWtPalAbsnt OR #s150_StChkNxtStRdyToRecvTTUp_T2 OR #s150_StChkNxtStRdyToRecvTTUp_T1 OR #s160_StWtFrStprDn_CnvyrStrt_T1) AND NOT #sStWtResetRel AND NOT #s165_StWtPalAbsnt_T1;
   IF #s165_StWtPalAbsnt THEN #StateNo := 165; END_IF;
END_REGION

REGION Network 62: Actions for STATE Num:165 StWtPalAbsnt
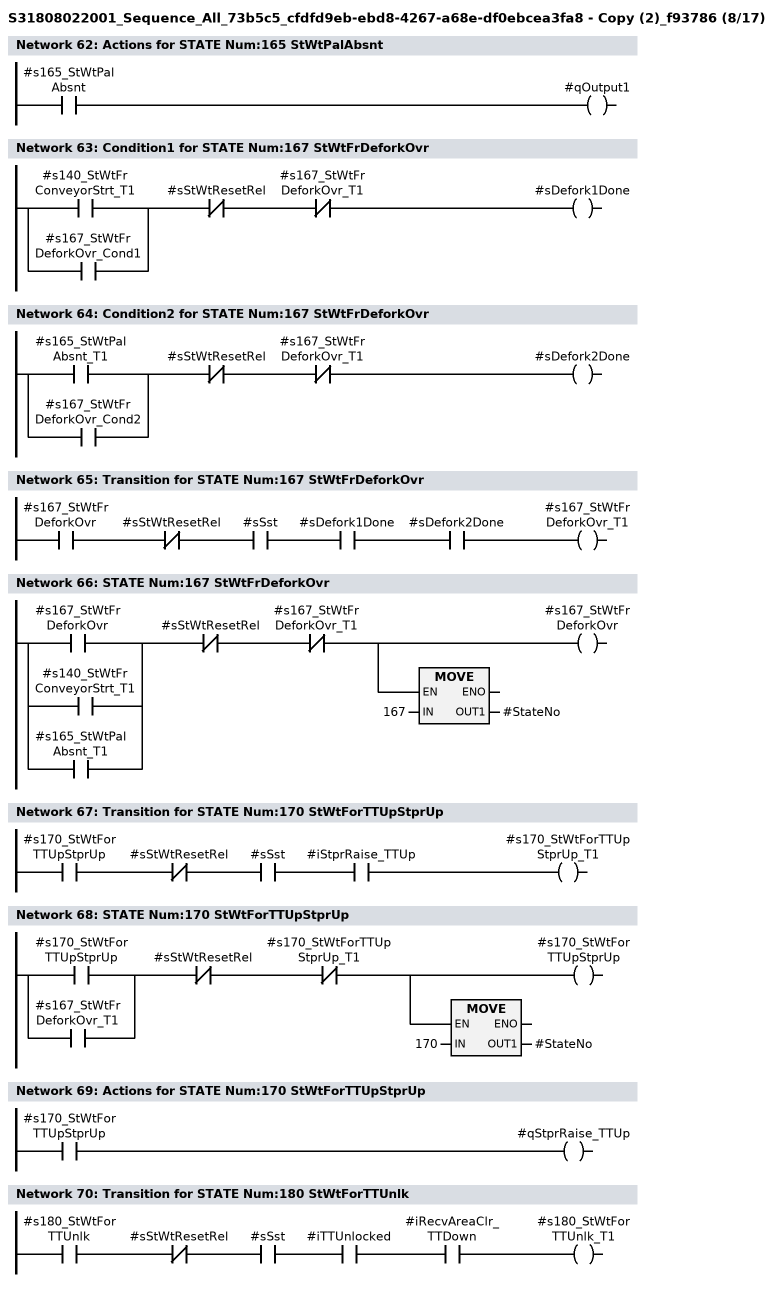
   RUNG wire#powerrail
      Contact( #s165_StWtPalAbsnt )
      Coil( #qOutput1 )
   END_RUNG
   // the same network as SCL:
   #qOutput1 := #s165_StWtPalAbsnt;
END_REGION

REGION Network 63: Condition1 for STATE Num:167 StWtFrDeforkOvr
   RUNG wire#powerrail
      Contact( #s140_StWtFrConveyorStrt_T1 )
      wire#w1
      I_Contact( #sStWtResetRel )
      I_Contact( #s167_StWtFrDeforkOvr_T1 )
      Coil( #sDefork1Done )
   END_RUNG
   RUNG wire#powerrail
      Contact( #s167_StWtFrDeforkOvr_Cond1 )
   END_RUNG wire#w1
   // the same network as SCL:
   #sDefork1Done := (#s140_StWtFrConveyorStrt_T1 OR #s167_StWtFrDeforkOvr_Cond1) AND NOT #sStWtResetRel AND NOT #s167_StWtFrDeforkOvr_T1;
END_REGION

REGION Network 64: Condition2 for STATE Num:167 StWtFrDeforkOvr
   RUNG wire#powerrail
      Contact( #s165_StWtPalAbsnt_T1 )
      wire#w1
      I_Contact( #sStWtResetRel )
      I_Contact( #s167_StWtFrDeforkOvr_T1 )
      Coil( #sDefork2Done )
   END_RUNG
   RUNG wire#powerrail
      Contact( #s167_StWtFrDeforkOvr_Cond2 )
   END_RUNG wire#w1
   // the same network as SCL:
   #sDefork2Done := (#s165_StWtPalAbsnt_T1 OR #s167_StWtFrDeforkOvr_Cond2) AND NOT #sStWtResetRel AND NOT #s167_StWtFrDeforkOvr_T1;
END_REGION

REGION Network 65: Transition for STATE Num:167 StWtFrDeforkOvr
   RUNG wire#powerrail
      Contact( #s167_StWtFrDeforkOvr )
      I_Contact( #sStWtResetRel )
      Contact( #sSst )
      Contact( #sDefork1Done )
      Contact( #sDefork2Done )
      Coil( #s167_StWtFrDeforkOvr_T1 )
   END_RUNG
   // the same network as SCL:
   #s167_StWtFrDeforkOvr_T1 := #s167_StWtFrDeforkOvr AND NOT #sStWtResetRel AND #sSst AND #sDefork1Done AND #sDefork2Done;
END_REGION

REGION Network 66: STATE Num:167 StWtFrDeforkOvr
   RUNG wire#powerrail
      Contact( #s167_StWtFrDeforkOvr )
      wire#w1
      I_Contact( #sStWtResetRel )
      I_Contact( #s167_StWtFrDeforkOvr_T1 )
      wire#w2
      Coil( #s167_StWtFrDeforkOvr )
   END_RUNG
   RUNG wire#powerrail
      Contact( #s140_StWtFrConveyorStrt_T1 )
   END_RUNG wire#w1
   RUNG wire#powerrail
      Contact( #s165_StWtPalAbsnt_T1 )
   END_RUNG wire#w1
   RUNG wire#w2
      { S7_GenerateENO := "TRUE" } Move(in := 167, out1 => #StateNo)
   END_RUNG
   // the same network as SCL:
   #s167_StWtFrDeforkOvr := (#s167_StWtFrDeforkOvr OR #s140_StWtFrConveyorStrt_T1 OR #s165_StWtPalAbsnt_T1) AND NOT #sStWtResetRel AND NOT #s167_StWtFrDeforkOvr_T1;
   IF #s167_StWtFrDeforkOvr THEN #StateNo := 167; END_IF;
END_REGION

REGION Network 67: Transition for STATE Num:170 StWtForTTUpStprUp
   RUNG wire#powerrail
      Contact( #s170_StWtForTTUpStprUp )
      I_Contact( #sStWtResetRel )
      Contact( #sSst )
      Contact( #iStprRaise_TTUp )
      Coil( #s170_StWtForTTUpStprUp_T1 )
   END_RUNG
   // the same network as SCL:
   #s170_StWtForTTUpStprUp_T1 := #s170_StWtForTTUpStprUp AND NOT #sStWtResetRel AND #sSst AND #iStprRaise_TTUp;
END_REGION

REGION Network 68: STATE Num:170 StWtForTTUpStprUp
   RUNG wire#powerrail
      Contact( #s170_StWtForTTUpStprUp )
      wire#w1
      I_Contact( #sStWtResetRel )
      I_Contact( #s170_StWtForTTUpStprUp_T1 )
      wire#w2
      Coil( #s170_StWtForTTUpStprUp )
   END_RUNG
   RUNG wire#powerrail
      Contact( #s167_StWtFrDeforkOvr_T1 )
   END_RUNG wire#w1
   RUNG wire#w2
      { S7_GenerateENO := "TRUE" } Move(in := 170, out1 => #StateNo)
   END_RUNG
   // the same network as SCL:
   #s170_StWtForTTUpStprUp := (#s170_StWtForTTUpStprUp OR #s167_StWtFrDeforkOvr_T1) AND NOT #sStWtResetRel AND NOT #s170_StWtForTTUpStprUp_T1;
   IF #s170_StWtForTTUpStprUp THEN #StateNo := 170; END_IF;
END_REGION

REGION Network 69: Actions for STATE Num:170 StWtForTTUpStprUp
   RUNG wire#powerrail
      Contact( #s170_StWtForTTUpStprUp )
      Coil( #qStprRaise_TTUp )
   END_RUNG
   // the same network as SCL:
   #qStprRaise_TTUp := #s170_StWtForTTUpStprUp;
END_REGION

REGION Network 70: Transition for STATE Num:180 StWtForTTUnlk
   RUNG wire#powerrail
      Contact( #s180_StWtForTTUnlk )
      I_Contact( #sStWtResetRel )
      Contact( #sSst )
      Contact( #iTTUnlocked )
      Contact( #iRecvAreaClr_TTDown )
      Coil( #s180_StWtForTTUnlk_T1 )
   END_RUNG
   // the same network as SCL:
   #s180_StWtForTTUnlk_T1 := #s180_StWtForTTUnlk AND NOT #sStWtResetRel AND #sSst AND #iTTUnlocked AND #iRecvAreaClr_TTDown;
END_REGION

REGION Network 71: STATE Num:180 StWtForTTUnlk
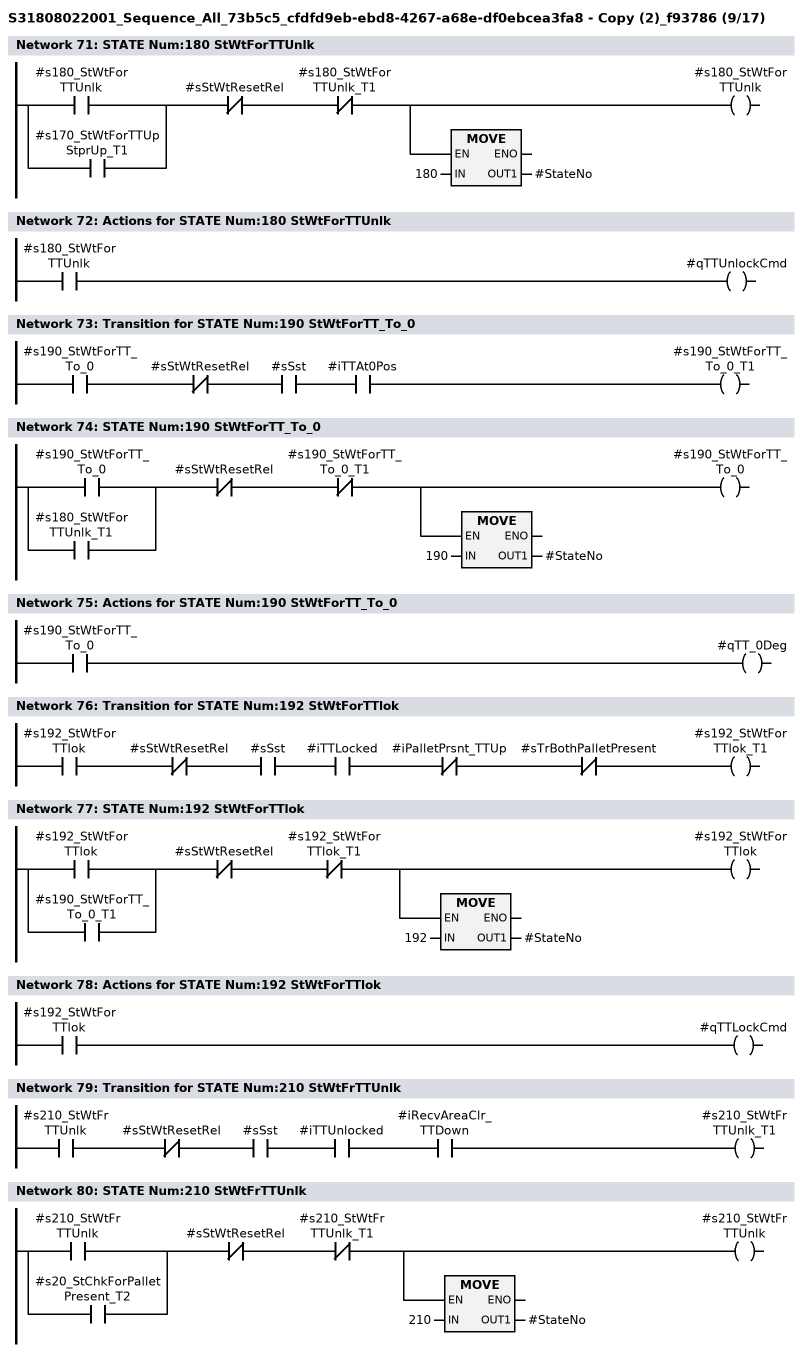
   RUNG wire#powerrail
      Contact( #s180_StWtForTTUnlk )
      wire#w1
      I_Contact( #sStWtResetRel )
      I_Contact( #s180_StWtForTTUnlk_T1 )
      wire#w2
      Coil( #s180_StWtForTTUnlk )
   END_RUNG
   RUNG wire#powerrail
      Contact( #s170_StWtForTTUpStprUp_T1 )
   END_RUNG wire#w1
   RUNG wire#w2
      { S7_GenerateENO := "TRUE" } Move(in := 180, out1 => #StateNo)
   END_RUNG
   // the same network as SCL:
   #s180_StWtForTTUnlk := (#s180_StWtForTTUnlk OR #s170_StWtForTTUpStprUp_T1) AND NOT #sStWtResetRel AND NOT #s180_StWtForTTUnlk_T1;
   IF #s180_StWtForTTUnlk THEN #StateNo := 180; END_IF;
END_REGION

REGION Network 72: Actions for STATE Num:180 StWtForTTUnlk
   RUNG wire#powerrail
      Contact( #s180_StWtForTTUnlk )
      Coil( #qTTUnlockCmd )
   END_RUNG
   // the same network as SCL:
   #qTTUnlockCmd := #s180_StWtForTTUnlk;
END_REGION

REGION Network 73: Transition for STATE Num:190 StWtForTT_To_0
   RUNG wire#powerrail
      Contact( #s190_StWtForTT_To_0 )
      I_Contact( #sStWtResetRel )
      Contact( #sSst )
      Contact( #iTTAt0Pos )
      Coil( #s190_StWtForTT_To_0_T1 )
   END_RUNG
   // the same network as SCL:
   #s190_StWtForTT_To_0_T1 := #s190_StWtForTT_To_0 AND NOT #sStWtResetRel AND #sSst AND #iTTAt0Pos;
END_REGION

REGION Network 74: STATE Num:190 StWtForTT_To_0
   RUNG wire#powerrail
      Contact( #s190_StWtForTT_To_0 )
      wire#w1
      I_Contact( #sStWtResetRel )
      I_Contact( #s190_StWtForTT_To_0_T1 )
      wire#w2
      Coil( #s190_StWtForTT_To_0 )
   END_RUNG
   RUNG wire#powerrail
      Contact( #s180_StWtForTTUnlk_T1 )
   END_RUNG wire#w1
   RUNG wire#w2
      { S7_GenerateENO := "TRUE" } Move(in := 190, out1 => #StateNo)
   END_RUNG
   // the same network as SCL:
   #s190_StWtForTT_To_0 := (#s190_StWtForTT_To_0 OR #s180_StWtForTTUnlk_T1) AND NOT #sStWtResetRel AND NOT #s190_StWtForTT_To_0_T1;
   IF #s190_StWtForTT_To_0 THEN #StateNo := 190; END_IF;
END_REGION

REGION Network 75: Actions for STATE Num:190 StWtForTT_To_0
   RUNG wire#powerrail
      Contact( #s190_StWtForTT_To_0 )
      Coil( #qTT_0Deg )
   END_RUNG
   // the same network as SCL:
   #qTT_0Deg := #s190_StWtForTT_To_0;
END_REGION

REGION Network 76: Transition for STATE Num:192 StWtForTTlok
   RUNG wire#powerrail
      Contact( #s192_StWtForTTlok )
      I_Contact( #sStWtResetRel )
      Contact( #sSst )
      Contact( #iTTLocked )
      I_Contact( #iPalletPrsnt_TTUp )
      I_Contact( #sTrBothPalletPresent )
      Coil( #s192_StWtForTTlok_T1 )
   END_RUNG
   // the same network as SCL:
   #s192_StWtForTTlok_T1 := #s192_StWtForTTlok AND NOT #sStWtResetRel AND #sSst AND #iTTLocked AND NOT #iPalletPrsnt_TTUp AND NOT #sTrBothPalletPresent;
END_REGION

REGION Network 77: STATE Num:192 StWtForTTlok
   RUNG wire#powerrail
      Contact( #s192_StWtForTTlok )
      wire#w1
      I_Contact( #sStWtResetRel )
      I_Contact( #s192_StWtForTTlok_T1 )
      wire#w2
      Coil( #s192_StWtForTTlok )
   END_RUNG
   RUNG wire#powerrail
      Contact( #s190_StWtForTT_To_0_T1 )
   END_RUNG wire#w1
   RUNG wire#w2
      { S7_GenerateENO := "TRUE" } Move(in := 192, out1 => #StateNo)
   END_RUNG
   // the same network as SCL:
   #s192_StWtForTTlok := (#s192_StWtForTTlok OR #s190_StWtForTT_To_0_T1) AND NOT #sStWtResetRel AND NOT #s192_StWtForTTlok_T1;
   IF #s192_StWtForTTlok THEN #StateNo := 192; END_IF;
END_REGION

REGION Network 78: Actions for STATE Num:192 StWtForTTlok
   RUNG wire#powerrail
      Contact( #s192_StWtForTTlok )
      Coil( #qTTLockCmd )
   END_RUNG
   // the same network as SCL:
   #qTTLockCmd := #s192_StWtForTTlok;
END_REGION

REGION Network 79: Transition for STATE Num:210 StWtFrTTUnlk
   RUNG wire#powerrail
      Contact( #s210_StWtFrTTUnlk )
      I_Contact( #sStWtResetRel )
      Contact( #sSst )
      Contact( #iTTUnlocked )
      Contact( #iRecvAreaClr_TTDown )
      Coil( #s210_StWtFrTTUnlk_T1 )
   END_RUNG
   // the same network as SCL:
   #s210_StWtFrTTUnlk_T1 := #s210_StWtFrTTUnlk AND NOT #sStWtResetRel AND #sSst AND #iTTUnlocked AND #iRecvAreaClr_TTDown;
END_REGION

REGION Network 80: STATE Num:210 StWtFrTTUnlk
   RUNG wire#powerrail
      Contact( #s210_StWtFrTTUnlk )
      wire#w1
      I_Contact( #sStWtResetRel )
      I_Contact( #s210_StWtFrTTUnlk_T1 )
      wire#w2
      Coil( #s210_StWtFrTTUnlk )
   END_RUNG
   RUNG wire#powerrail
      Contact( #s20_StChkForPalletPresent_T2 )
   END_RUNG wire#w1
   RUNG wire#w2
      { S7_GenerateENO := "TRUE" } Move(in := 210, out1 => #StateNo)
   END_RUNG
   // the same network as SCL:
   #s210_StWtFrTTUnlk := (#s210_StWtFrTTUnlk OR #s20_StChkForPalletPresent_T2) AND NOT #sStWtResetRel AND NOT #s210_StWtFrTTUnlk_T1;
   IF #s210_StWtFrTTUnlk THEN #StateNo := 210; END_IF;
END_REGION

REGION Network 81: Actions for STATE Num:210 StWtFrTTUnlk
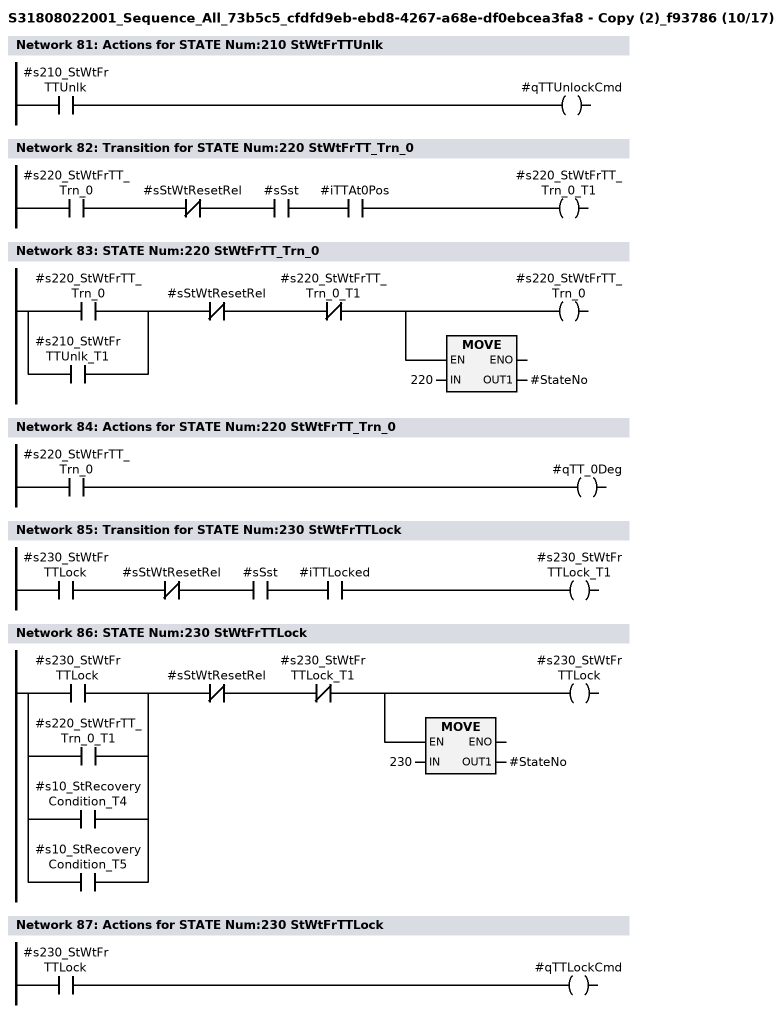
   RUNG wire#powerrail
      Contact( #s210_StWtFrTTUnlk )
      Coil( #qTTUnlockCmd )
   END_RUNG
   // the same network as SCL:
   #qTTUnlockCmd := #s210_StWtFrTTUnlk;
END_REGION

REGION Network 82: Transition for STATE Num:220 StWtFrTT_Trn_0
   RUNG wire#powerrail
      Contact( #s220_StWtFrTT_Trn_0 )
      I_Contact( #sStWtResetRel )
      Contact( #sSst )
      Contact( #iTTAt0Pos )
      Coil( #s220_StWtFrTT_Trn_0_T1 )
   END_RUNG
   // the same network as SCL:
   #s220_StWtFrTT_Trn_0_T1 := #s220_StWtFrTT_Trn_0 AND NOT #sStWtResetRel AND #sSst AND #iTTAt0Pos;
END_REGION

REGION Network 83: STATE Num:220 StWtFrTT_Trn_0
   RUNG wire#powerrail
      Contact( #s220_StWtFrTT_Trn_0 )
      wire#w1
      I_Contact( #sStWtResetRel )
      I_Contact( #s220_StWtFrTT_Trn_0_T1 )
      wire#w2
      Coil( #s220_StWtFrTT_Trn_0 )
   END_RUNG
   RUNG wire#powerrail
      Contact( #s210_StWtFrTTUnlk_T1 )
   END_RUNG wire#w1
   RUNG wire#w2
      { S7_GenerateENO := "TRUE" } Move(in := 220, out1 => #StateNo)
   END_RUNG
   // the same network as SCL:
   #s220_StWtFrTT_Trn_0 := (#s220_StWtFrTT_Trn_0 OR #s210_StWtFrTTUnlk_T1) AND NOT #sStWtResetRel AND NOT #s220_StWtFrTT_Trn_0_T1;
   IF #s220_StWtFrTT_Trn_0 THEN #StateNo := 220; END_IF;
END_REGION

REGION Network 84: Actions for STATE Num:220 StWtFrTT_Trn_0
   RUNG wire#powerrail
      Contact( #s220_StWtFrTT_Trn_0 )
      Coil( #qTT_0Deg )
   END_RUNG
   // the same network as SCL:
   #qTT_0Deg := #s220_StWtFrTT_Trn_0;
END_REGION

REGION Network 85: Transition for STATE Num:230 StWtFrTTLock
   RUNG wire#powerrail
      Contact( #s230_StWtFrTTLock )
      I_Contact( #sStWtResetRel )
      Contact( #sSst )
      Contact( #iTTLocked )
      Coil( #s230_StWtFrTTLock_T1 )
   END_RUNG
   // the same network as SCL:
   #s230_StWtFrTTLock_T1 := #s230_StWtFrTTLock AND NOT #sStWtResetRel AND #sSst AND #iTTLocked;
END_REGION

REGION Network 86: STATE Num:230 StWtFrTTLock
   RUNG wire#powerrail
      Contact( #s230_StWtFrTTLock )
      wire#w1
      I_Contact( #sStWtResetRel )
      I_Contact( #s230_StWtFrTTLock_T1 )
      wire#w2
      Coil( #s230_StWtFrTTLock )
   END_RUNG
   RUNG wire#powerrail
      Contact( #s220_StWtFrTT_Trn_0_T1 )
   END_RUNG wire#w1
   RUNG wire#powerrail
      Contact( #s10_StRecoveryCondition_T4 )
   END_RUNG wire#w1
   RUNG wire#powerrail
      Contact( #s10_StRecoveryCondition_T5 )
   END_RUNG wire#w1
   RUNG wire#w2
      { S7_GenerateENO := "TRUE" } Move(in := 230, out1 => #StateNo)
   END_RUNG
   // the same network as SCL:
   #s230_StWtFrTTLock := (#s230_StWtFrTTLock OR #s220_StWtFrTT_Trn_0_T1 OR #s10_StRecoveryCondition_T4 OR #s10_StRecoveryCondition_T5) AND NOT #sStWtResetRel AND NOT #s230_StWtFrTTLock_T1;
   IF #s230_StWtFrTTLock THEN #StateNo := 230; END_IF;
END_REGION

REGION Network 87: Actions for STATE Num:230 StWtFrTTLock
   RUNG wire#powerrail
      Contact( #s230_StWtFrTTLock )
      Coil( #qTTLockCmd )
   END_RUNG
   // the same network as SCL:
   #qTTLockCmd := #s230_StWtFrTTLock;
END_REGION

